ABB RAPID module: Ingenieria165.mod

MODULE Ingenieria165
    !***********************************************************
    !
    ! Modulo:  Ingenieria165
    !
    ! Descripción:
    !   Modulo con rutinas para decoracion con el motivo 165 años de facultad de ingeneria
    !
    ! Autor: Juan_Daleman
    !
    ! Versión: 1.0
    !
    !***********************************************************
    CONST robtarget Target_Tap165_10:=[[81.313,-88.677,-19.266],[0.707106781,0,0,0.707106781],[0,0,0,0],[9E+09,9E+09,9E+09,9E+09,9E+09,9E+09]];
    CONST robtarget Target_Tap165_20:=[[81.313,-88.677,-2.266],[0.707106781,0,0,0.707106781],[0,0,0,0],[9E+09,9E+09,9E+09,9E+09,9E+09,9E+09]];
    CONST robtarget Target_Tap165_30:=[[81.338,-82.631,-2.266],[0.707106781,0,0,0.707106781],[0,0,0,0],[9E+09,9E+09,9E+09,9E+09,9E+09,9E+09]];
    CONST robtarget Target_Tap165_40:=[[76.897,-82.904,-2.306],[0.707106781,0,0,0.707106781],[0,0,0,0],[9E+09,9E+09,9E+09,9E+09,9E+09,9E+09]];
    CONST robtarget Target_Tap165_50:=[[81.369,-82.46,-2.266],[0.707106781,0,0,0.707106781],[0,0,0,0],[9E+09,9E+09,9E+09,9E+09,9E+09,9E+09]];
    CONST robtarget Target_Tap165_60:=[[81.524,-77.183,-2.264],[0.707106781,0,0,0.707106781],[0,0,0,0],[9E+09,9E+09,9E+09,9E+09,9E+09,9E+09]];
    CONST robtarget Target_Tap165_70:=[[75.87,-77.461,-2.316],[0.707106781,0,0,0.707106781],[0,0,0,0],[9E+09,9E+09,9E+09,9E+09,9E+09,9E+09]];
    CONST robtarget Target_Tap165_80:=[[75.87,-77.461,-20],[0.707106781,0,0,0.707106781],[0,0,0,0],[9E+09,9E+09,9E+09,9E+09,9E+09,9E+09]];
    CONST robtarget Target_Tap165_90:=[[67.923,-79.66,-20],[0.707106781,0,0,0.707106781],[0,0,0,0],[9E+09,9E+09,9E+09,9E+09,9E+09,9E+09]];
    CONST robtarget Target_Tap165_100:=[[67.923,-79.66,-2.388],[0.707106781,0,0,0.707106781],[0,0,0,0],[9E+09,9E+09,9E+09,9E+09,9E+09,9E+09]];
    CONST robtarget Target_Tap165_110:=[[67.877,-88.682,-2.388],[0.707106781,0,0,0.707106781],[0,0,0,0],[9E+09,9E+09,9E+09,9E+09,9E+09,9E+09]];
    CONST robtarget Target_Tap165_120:=[[69.176,-87.545,-2.376],[0.707106781,0,0,0.707106781],[0,0,0,0],[9E+09,9E+09,9E+09,9E+09,9E+09,9E+09]];
    CONST robtarget Target_Tap165_130:=[[73.466,-88.301,-2.338],[0.707106781,0,0,0.707106781],[0,0,0,0],[9E+09,9E+09,9E+09,9E+09,9E+09,9E+09]];
    CONST robtarget Target_Tap165_140:=[[75.281,-84.884,-2.321],[0.707106781,0,0,0.707106781],[0,0,0,0],[9E+09,9E+09,9E+09,9E+09,9E+09,9E+09]];
    CONST robtarget Target_Tap165_150:=[[72.745,-79.717,-2.344],[0.707106781,0,0,0.707106781],[0,0,0,0],[9E+09,9E+09,9E+09,9E+09,9E+09,9E+09]];
    CONST robtarget Target_Tap165_160:=[[69.243,-80.87,-2.376],[0.707106781,0,0,0.707106781],[0,0,0,0],[9E+09,9E+09,9E+09,9E+09,9E+09,9E+09]];
    CONST robtarget Target_Tap165_170:=[[69.243,-80.87,-20],[0.707106781,0,0,0.707106781],[0,0,0,0],[9E+09,9E+09,9E+09,9E+09,9E+09,9E+09]];
    CONST robtarget Target_Tap165_180:=[[57.703,-85.818,-20],[0.707106781,0,0,0.707106781],[0,0,0,0],[9E+09,9E+09,9E+09,9E+09,9E+09,9E+09]];
    CONST robtarget Target_Tap165_190:=[[57.683,-85.747,-2.481],[0.707106781,0,0,0.707106781],[0,0,0,0],[9E+09,9E+09,9E+09,9E+09,9E+09,9E+09]];
    CONST robtarget Target_Tap165_200:=[[62.028,-88.896,-2.441],[0.707106781,0,0,0.707106781],[0,0,0,0],[9E+09,9E+09,9E+09,9E+09,9E+09,9E+09]];
    CONST robtarget Target_Tap165_210:=[[65.482,-83.568,-2.41],[0.707106781,0,0,0.707106781],[0,0,0,0],[9E+09,9E+09,9E+09,9E+09,9E+09,9E+09]];
    CONST robtarget Target_Tap165_220:=[[61.822,-79.686,-2.443],[0.707106781,0,0,0.707106781],[0,0,0,0],[9E+09,9E+09,9E+09,9E+09,9E+09,9E+09]];
    CONST robtarget Target_Tap165_230:=[[57.626,-82.905,-2.481],[0.707106781,0,0,0.707106781],[0,0,0,0],[9E+09,9E+09,9E+09,9E+09,9E+09,9E+09]];
    CONST robtarget Target_Tap165_240:=[[57.626,-82.905,-20],[0.707106781,0,0,0.707106781],[0,0,0,0],[9E+09,9E+09,9E+09,9E+09,9E+09,9E+09]];
    CONST robtarget Target_Tap165_250:=[[55.482,-79.946,-20],[0.707106781,0,0,0.707106781],[0,0,0,0],[9E+09,9E+09,9E+09,9E+09,9E+09,9E+09]];
    CONST robtarget Target_Tap165_260:=[[55.542,-79.789,-2.5],[0.707106781,0,0,0.707106781],[0,0,0,0],[9E+09,9E+09,9E+09,9E+09,9E+09,9E+09]];
    CONST robtarget Target_Tap165_270:=[[55.414,-88.257,-2.501],[0.707106781,0,0,0.707106781],[0,0,0,0],[9E+09,9E+09,9E+09,9E+09,9E+09,9E+09]];
    CONST robtarget Target_Tap165_280:=[[53.088,-88.957,-2.522],[0.707106781,0,0,0.707106781],[0,0,0,0],[9E+09,9E+09,9E+09,9E+09,9E+09,9E+09]];
    CONST robtarget Target_Tap165_290:=[[50.869,-87.673,-2.542],[0.707106781,0,0,0.707106781],[0,0,0,0],[9E+09,9E+09,9E+09,9E+09,9E+09,9E+09]];
    CONST robtarget Target_Tap165_300:=[[49.455,-88.876,-2.555],[0.707106781,0,0,0.707106781],[0,0,0,0],[9E+09,9E+09,9E+09,9E+09,9E+09,9E+09]];
    CONST robtarget Target_Tap165_310:=[[49.666,-79.854,-2.553],[0.707106781,0,0,0.707106781],[0,0,0,0],[9E+09,9E+09,9E+09,9E+09,9E+09,9E+09]];
    CONST robtarget Target_Tap165_320:=[[49.666,-79.854,-20],[0.707106781,0,0,0.707106781],[0,0,0,0],[9E+09,9E+09,9E+09,9E+09,9E+09,9E+09]];
    CONST robtarget Target_Tap165_330:=[[45.617,-88.918,-20],[0.707106781,0,0,0.707106781],[0,0,0,0],[9E+09,9E+09,9E+09,9E+09,9E+09,9E+09]];
    CONST robtarget Target_Tap165_340:=[[45.617,-88.918,-2.59],[0.707106781,0,0,0.707106781],[0,0,0,0],[9E+09,9E+09,9E+09,9E+09,9E+09,9E+09]];
    CONST robtarget Target_Tap165_350:=[[45.551,-76.897,-2.591],[0.707106781,0,0,0.707106781],[0,0,0,0],[9E+09,9E+09,9E+09,9E+09,9E+09,9E+09]];
    CONST robtarget Target_Tap165_360:=[[45.551,-76.897,-23],[0.707106781,0,0,0.707106781],[0,0,0,0],[9E+09,9E+09,9E+09,9E+09,9E+09,9E+09]];
    CONST robtarget Target_Tap165_370:=[[41.407,-77.76,-20],[0.707106781,0,0,0.707106781],[0,0,0,0],[9E+09,9E+09,9E+09,9E+09,9E+09,9E+09]];
    CONST robtarget Target_Tap165_380:=[[41.407,-77.76,0.372],[0.707106781,0,0,0.707106781],[0,0,0,0],[9E+09,9E+09,9E+09,9E+09,9E+09,9E+09]];
    CONST robtarget Target_Tap165_390:=[[41.282,-80.994,-2.629],[0.707106781,0,0,0.707106781],[0,0,0,0],[9E+09,9E+09,9E+09,9E+09,9E+09,9E+09]];
    CONST robtarget Target_Tap165_400:=[[43.422,-80.77,-2.61],[0.707106781,0,0,0.707106781],[0,0,0,0],[9E+09,9E+09,9E+09,9E+09,9E+09,9E+09]];
    CONST robtarget Target_Tap165_410:=[[38.361,-80.952,-2.656],[0.707106781,0,0,0.707106781],[0,0,0,0],[9E+09,9E+09,9E+09,9E+09,9E+09,9E+09]];
    CONST robtarget Target_Tap165_420:=[[41.333,-81.008,-2.629],[0.707106781,0,0,0.707106781],[0,0,0,0],[9E+09,9E+09,9E+09,9E+09,9E+09,9E+09]];
    CONST robtarget Target_Tap165_430:=[[41.267,-88.487,-2.629],[0.707106781,0,0,0.707106781],[0,0,0,0],[9E+09,9E+09,9E+09,9E+09,9E+09,9E+09]];
    CONST robtarget Target_Tap165_440:=[[38.45,-88.997,-2.655],[0.707106781,0,0,0.707106781],[0,0,0,0],[9E+09,9E+09,9E+09,9E+09,9E+09,9E+09]];
    CONST robtarget Target_Tap165_450:=[[38.45,-88.997,-20],[0.707106781,0,0,0.707106781],[0,0,0,0],[9E+09,9E+09,9E+09,9E+09,9E+09,9E+09]];
    CONST robtarget Target_Tap165_460:=[[30.389,-80.073,-20],[0.707106781,0,0,0.707106781],[0,0,0,0],[9E+09,9E+09,9E+09,9E+09,9E+09,9E+09]];
    CONST robtarget Target_Tap165_470:=[[30.389,-80.073,-2.728],[0.707106781,0,0,0.707106781],[0,0,0,0],[9E+09,9E+09,9E+09,9E+09,9E+09,9E+09]];
    CONST robtarget Target_Tap165_480:=[[30.235,-89.097,-2.73],[0.707106781,0,0,0.707106781],[0,0,0,0],[9E+09,9E+09,9E+09,9E+09,9E+09,9E+09]];
    CONST robtarget Target_Tap165_490:=[[31.518,-87.896,-2.718],[0.707106781,0,0,0.707106781],[0,0,0,0],[9E+09,9E+09,9E+09,9E+09,9E+09,9E+09]];
    CONST robtarget Target_Tap165_500:=[[34.632,-89.19,-2.69],[0.707106781,0,0,0.707106781],[0,0,0,0],[9E+09,9E+09,9E+09,9E+09,9E+09,9E+09]];
    CONST robtarget Target_Tap165_510:=[[37.622,-85.047,-2.663],[0.707106781,0,0,0.707106781],[0,0,0,0],[9E+09,9E+09,9E+09,9E+09,9E+09,9E+09]];
    CONST robtarget Target_Tap165_520:=[[35.565,-79.921,-2.682],[0.707106781,0,0,0.707106781],[0,0,0,0],[9E+09,9E+09,9E+09,9E+09,9E+09,9E+09]];
    CONST robtarget Target_Tap165_530:=[[31.419,-81.282,-2.719],[0.707106781,0,0,0.707106781],[0,0,0,0],[9E+09,9E+09,9E+09,9E+09,9E+09,9E+09]];
    CONST robtarget Target_Tap165_540:=[[31.419,-81.282,-20],[0.707106781,0,0,0.707106781],[0,0,0,0],[9E+09,9E+09,9E+09,9E+09,9E+09,9E+09]];
    CONST robtarget Target_Tap165_550:=[[20.747,-77.17,-20],[0.707106781,0,0,0.707106781],[0,0,0,0],[9E+09,9E+09,9E+09,9E+09,9E+09,9E+09]];
    CONST robtarget Target_Tap165_560:=[[20.805,-77.169,-2.815],[0.707106781,0,0,0.707106781],[0,0,0,0],[9E+09,9E+09,9E+09,9E+09,9E+09,9E+09]];
    CONST robtarget Target_Tap165_570:=[[20.61,-89.193,-2.817],[0.707106781,0,0,0.707106781],[0,0,0,0],[9E+09,9E+09,9E+09,9E+09,9E+09,9E+09]];
    CONST robtarget Target_Tap165_580:=[[21.819,-88.233,-2.806],[0.707106781,0,0,0.707106781],[0,0,0,0],[9E+09,9E+09,9E+09,9E+09,9E+09,9E+09]];
    CONST robtarget Target_Tap165_590:=[[25.21,-89.217,-2.775],[0.707106781,0,0,0.707106781],[0,0,0,0],[9E+09,9E+09,9E+09,9E+09,9E+09,9E+09]];
    CONST robtarget Target_Tap165_600:=[[27.949,-85.408,-2.75],[0.707106781,0,0,0.707106781],[0,0,0,0],[9E+09,9E+09,9E+09,9E+09,9E+09,9E+09]];
    CONST robtarget Target_Tap165_610:=[[25.874,-80.415,-2.769],[0.707106781,0,0,0.707106781],[0,0,0,0],[9E+09,9E+09,9E+09,9E+09,9E+09,9E+09]];
    CONST robtarget Target_Tap165_620:=[[21.748,-81.419,-2.807],[0.707106781,0,0,0.707106781],[0,0,0,0],[9E+09,9E+09,9E+09,9E+09,9E+09,9E+09]];
    CONST robtarget Target_Tap165_630:=[[21.748,-81.419,-20],[0.707106781,0,0,0.707106781],[0,0,0,0],[9E+09,9E+09,9E+09,9E+09,9E+09,9E+09]];
    CONST robtarget Target_Tap165_640:=[[8.35,-77.306,-20],[0.707106781,0,0,0.707106781],[0,0,0,0],[9E+09,9E+09,9E+09,9E+09,9E+09,9E+09]];
    CONST robtarget Target_Tap165_650:=[[8.35,-77.306,-2.928],[0.707106781,0,0,0.707106781],[0,0,0,0],[9E+09,9E+09,9E+09,9E+09,9E+09,9E+09]];
    CONST robtarget Target_Tap165_660:=[[7.975,-89.332,-2.932],[0.707106781,0,0,0.707106781],[0,0,0,0],[9E+09,9E+09,9E+09,9E+09,9E+09,9E+09]];
    CONST robtarget Target_Tap165_670:=[[9.494,-88.106,-2.918],[0.707106781,0,0,0.707106781],[0,0,0,0],[9E+09,9E+09,9E+09,9E+09,9E+09,9E+09]];
    CONST robtarget Target_Tap165_680:=[[13.081,-89.294,-2.885],[0.707106781,0,0,0.707106781],[0,0,0,0],[9E+09,9E+09,9E+09,9E+09,9E+09,9E+09]];
    CONST robtarget Target_Tap165_690:=[[15.593,-85.146,-2.863],[0.707106781,0,0,0.707106781],[0,0,0,0],[9E+09,9E+09,9E+09,9E+09,9E+09,9E+09]];
    CONST robtarget Target_Tap165_700:=[[13.446,-80.526,-2.882],[0.707106781,0,0,0.707106781],[0,0,0,0],[9E+09,9E+09,9E+09,9E+09,9E+09,9E+09]];
    CONST robtarget Target_Tap165_710:=[[9.38,-81.539,-2.919],[0.707106781,0,0,0.707106781],[0,0,0,0],[9E+09,9E+09,9E+09,9E+09,9E+09,9E+09]];
    CONST robtarget Target_Tap165_720:=[[9.38,-81.539,-20],[0.707106781,0,0,0.707106781],[0,0,0,0],[9E+09,9E+09,9E+09,9E+09,9E+09,9E+09]];
    CONST robtarget Target_Tap165_730:=[[-2.035,-86.612,-20],[0.707106781,0,0,0.707106781],[0,0,0,0],[9E+09,9E+09,9E+09,9E+09,9E+09,9E+09]];
    CONST robtarget Target_Tap165_740:=[[-2.035,-86.612,-3.023],[0.707106781,0,0,0.707106781],[0,0,0,0],[9E+09,9E+09,9E+09,9E+09,9E+09,9E+09]];
    CONST robtarget Target_Tap165_750:=[[2.246,-89.541,-2.984],[0.707106781,0,0,0.707106781],[0,0,0,0],[9E+09,9E+09,9E+09,9E+09,9E+09,9E+09]];
    CONST robtarget Target_Tap165_760:=[[5.81,-84.927,-2.951],[0.707106781,0,0,0.707106781],[0,0,0,0],[9E+09,9E+09,9E+09,9E+09,9E+09,9E+09]];
    CONST robtarget Target_Tap165_770:=[[1.692,-80.318,-2.989],[0.707106781,0,0,0.707106781],[0,0,0,0],[9E+09,9E+09,9E+09,9E+09,9E+09,9E+09]];
    CONST robtarget Target_Tap165_780:=[[-2.242,-85.619,-3.024],[0.707106781,0,0,0.707106781],[0,0,0,0],[9E+09,9E+09,9E+09,9E+09,9E+09,9E+09]];
    CONST robtarget Target_Tap165_790:=[[3.474,-85.692,-2.973],[0.707106781,0,0,0.707106781],[0,0,0,0],[9E+09,9E+09,9E+09,9E+09,9E+09,9E+09]];
    CONST robtarget Target_Tap165_800:=[[3.474,-85.692,-20],[0.707106781,0,0,0.707106781],[0,0,0,0],[9E+09,9E+09,9E+09,9E+09,9E+09,9E+09]];
    CONST robtarget Target_Tap165_810:=[[-7.455,-89.529,-20],[0.707106781,0,0,0.707106781],[0,0,0,0],[9E+09,9E+09,9E+09,9E+09,9E+09,9E+09]];
    CONST robtarget Target_Tap165_820:=[[-7.455,-89.529,-3.072],[0.707106781,0,0,0.707106781],[0,0,0,0],[9E+09,9E+09,9E+09,9E+09,9E+09,9E+09]];
    CONST robtarget Target_Tap165_830:=[[-7.408,-78.16,-3.071],[0.707106781,0,0,0.707106781],[0,0,0,0],[9E+09,9E+09,9E+09,9E+09,9E+09,9E+09]];
    CONST robtarget Target_Tap165_840:=[[-7.408,-78.16,-20],[0.707106781,0,0,0.707106781],[0,0,0,0],[9E+09,9E+09,9E+09,9E+09,9E+09,9E+09]];
    CONST robtarget Target_Tap165_850:=[[-11.373,-89.538,-20],[0.707106781,0,0,0.707106781],[0,0,0,0],[9E+09,9E+09,9E+09,9E+09,9E+09,9E+09]];
    CONST robtarget Target_Tap165_860:=[[-11.373,-89.538,-3.107],[0.707106781,0,0,0.707106781],[0,0,0,0],[9E+09,9E+09,9E+09,9E+09,9E+09,9E+09]];
    CONST robtarget Target_Tap165_870:=[[-11.145,-80.51,-3.105],[0.707106781,0,0,0.707106781],[0,0,0,0],[9E+09,9E+09,9E+09,9E+09,9E+09,9E+09]];
    CONST robtarget Target_Tap165_880:=[[-12.596,-81.788,-3.118],[0.707106781,0,0,0.707106781],[0,0,0,0],[9E+09,9E+09,9E+09,9E+09,9E+09,9E+09]];
    CONST robtarget Target_Tap165_890:=[[-15.49,-80.547,-3.145],[0.707106781,0,0,0.707106781],[0,0,0,0],[9E+09,9E+09,9E+09,9E+09,9E+09,9E+09]];
    CONST robtarget Target_Tap165_900:=[[-18.209,-83.364,-3.169],[0.707106781,0,0,0.707106781],[0,0,0,0],[9E+09,9E+09,9E+09,9E+09,9E+09,9E+09]];
    CONST robtarget Target_Tap165_910:=[[-18.164,-89.619,-3.169],[0.707106781,0,0,0.707106781],[0,0,0,0],[9E+09,9E+09,9E+09,9E+09,9E+09,9E+09]];
    CONST robtarget Target_Tap165_920:=[[-18.164,-89.619,-20],[0.707106781,0,0,0.707106781],[0,0,0,0],[9E+09,9E+09,9E+09,9E+09,9E+09,9E+09]];
    CONST robtarget Target_Tap165_930:=[[-19.664,-90.875,-20],[0.707106781,0,0,0.707106781],[0,0,0,0],[9E+09,9E+09,9E+09,9E+09,9E+09,9E+09]];
    CONST robtarget Target_Tap165_940:=[[-19.664,-90.875,-3.183],[0.707106781,0,0,0.707106781],[0,0,0,0],[9E+09,9E+09,9E+09,9E+09,9E+09,9E+09]];
    CONST robtarget Target_Tap165_950:=[[-24.113,-94.259,-3.223],[0.707106781,0,0,0.707106781],[0,0,0,0],[9E+09,9E+09,9E+09,9E+09,9E+09,9E+09]];
    CONST robtarget Target_Tap165_960:=[[-27.791,-90.884,-3.256],[0.707106781,0,0,0.707106781],[0,0,0,0],[9E+09,9E+09,9E+09,9E+09,9E+09,9E+09]];
    CONST robtarget Target_Tap165_970:=[[-27.929,-80.7,-3.258],[0.707106781,0,0,0.707106781],[0,0,0,0],[9E+09,9E+09,9E+09,9E+09,9E+09,9E+09]];
    CONST robtarget Target_Tap165_980:=[[-25.441,-81.899,-3.235],[0.707106781,0,0,0.707106781],[0,0,0,0],[9E+09,9E+09,9E+09,9E+09,9E+09,9E+09]];
    CONST robtarget Target_Tap165_990:=[[-22.502,-80.601,-3.208],[0.707106781,0,0,0.707106781],[0,0,0,0],[9E+09,9E+09,9E+09,9E+09,9E+09,9E+09]];
    CONST robtarget Target_Tap165_1000:=[[-19.387,-85.991,-3.18],[0.707106781,0,0,0.707106781],[0,0,0,0],[9E+09,9E+09,9E+09,9E+09,9E+09,9E+09]];
    CONST robtarget Target_Tap165_1010:=[[-21.158,-89.313,-3.196],[0.707106781,0,0,0.707106781],[0,0,0,0],[9E+09,9E+09,9E+09,9E+09,9E+09,9E+09]];
    CONST robtarget Target_Tap165_1020:=[[-25.481,-88.527,-3.235],[0.707106781,0,0,0.707106781],[0,0,0,0],[9E+09,9E+09,9E+09,9E+09,9E+09,9E+09]];
    CONST robtarget Target_Tap165_1030:=[[-25.431,-88.495,-20],[0.707106781,0,0,0.707106781],[0,0,0,0],[9E+09,9E+09,9E+09,9E+09,9E+09,9E+09]];
    CONST robtarget Target_Tap165_1040:=[[-36.83,-87.065,-20],[0.707106781,0,0,0.707106781],[0,0,0,0],[9E+09,9E+09,9E+09,9E+09,9E+09,9E+09]];
    CONST robtarget Target_Tap165_1050:=[[-36.83,-87.065,-3.338],[0.707106781,0,0,0.707106781],[0,0,0,0],[9E+09,9E+09,9E+09,9E+09,9E+09,9E+09]];
    CONST robtarget Target_Tap165_1060:=[[-32.555,-89.922,-3.3],[0.707106781,0,0,0.707106781],[0,0,0,0],[9E+09,9E+09,9E+09,9E+09,9E+09,9E+09]];
    CONST robtarget Target_Tap165_1070:=[[-29.008,-85.405,-3.267],[0.707106781,0,0,0.707106781],[0,0,0,0],[9E+09,9E+09,9E+09,9E+09,9E+09,9E+09]];
    CONST robtarget Target_Tap165_1080:=[[-33.253,-80.703,-3.306],[0.707106781,0,0,0.707106781],[0,0,0,0],[9E+09,9E+09,9E+09,9E+09,9E+09,9E+09]];
    CONST robtarget Target_Tap165_1090:=[[-37.045,-86.192,-3.34],[0.707106781,0,0,0.707106781],[0,0,0,0],[9E+09,9E+09,9E+09,9E+09,9E+09,9E+09]];
    CONST robtarget Target_Tap165_1100:=[[-31.341,-85.939,-3.289],[0.707106781,0,0,0.707106781],[0,0,0,0],[9E+09,9E+09,9E+09,9E+09,9E+09,9E+09]];
    CONST robtarget Target_Tap165_1110:=[[-31.341,-85.939,-20],[0.707106781,0,0,0.707106781],[0,0,0,0],[9E+09,9E+09,9E+09,9E+09,9E+09,9E+09]];
    CONST robtarget Target_Tap165_1120:=[[-39.521,-89.847,-20],[0.707106781,0,0,0.707106781],[0,0,0,0],[9E+09,9E+09,9E+09,9E+09,9E+09,9E+09]];
    CONST robtarget Target_Tap165_1130:=[[-39.521,-89.847,-3.363],[0.707106781,0,0,0.707106781],[0,0,0,0],[9E+09,9E+09,9E+09,9E+09,9E+09,9E+09]];
    CONST robtarget Target_Tap165_1140:=[[-39.341,-80.799,-3.361],[0.707106781,0,0,0.707106781],[0,0,0,0],[9E+09,9E+09,9E+09,9E+09,9E+09,9E+09]];
    CONST robtarget Target_Tap165_1150:=[[-40.79,-82.023,-3.374],[0.707106781,0,0,0.707106781],[0,0,0,0],[9E+09,9E+09,9E+09,9E+09,9E+09,9E+09]];
    CONST robtarget Target_Tap165_1160:=[[-43.877,-80.891,-3.402],[0.707106781,0,0,0.707106781],[0,0,0,0],[9E+09,9E+09,9E+09,9E+09,9E+09,9E+09]];
    CONST robtarget Target_Tap165_1170:=[[-46.356,-83.847,-3.425],[0.707106781,0,0,0.707106781],[0,0,0,0],[9E+09,9E+09,9E+09,9E+09,9E+09,9E+09]];
    CONST robtarget Target_Tap165_1180:=[[-46.289,-89.929,-3.424],[0.707106781,0,0,0.707106781],[0,0,0,0],[9E+09,9E+09,9E+09,9E+09,9E+09,9E+09]];
    CONST robtarget Target_Tap165_1190:=[[-46.289,-89.929,-20],[0.707106781,0,0,0.707106781],[0,0,0,0],[9E+09,9E+09,9E+09,9E+09,9E+09,9E+09]];
    CONST robtarget Target_Tap165_1200:=[[-49.014,-89.958,-20],[0.707106781,0,0,0.707106781],[0,0,0,0],[9E+09,9E+09,9E+09,9E+09,9E+09,9E+09]];
    CONST robtarget Target_Tap165_1210:=[[-49.014,-89.958,-3.449],[0.707106781,0,0,0.707106781],[0,0,0,0],[9E+09,9E+09,9E+09,9E+09,9E+09,9E+09]];
    CONST robtarget Target_Tap165_1220:=[[-48.979,-81.092,-3.449],[0.707106781,0,0,0.707106781],[0,0,0,0],[9E+09,9E+09,9E+09,9E+09,9E+09,9E+09]];
    CONST robtarget Target_Tap165_1230:=[[-48.979,-81.092,-20],[0.707106781,0,0,0.707106781],[0,0,0,0],[9E+09,9E+09,9E+09,9E+09,9E+09,9E+09]];
    CONST robtarget Target_Tap165_1240:=[[-49.066,-76.978,-20],[0.707106781,0,0,0.707106781],[0,0,0,0],[9E+09,9E+09,9E+09,9E+09,9E+09,9E+09]];
    CONST robtarget Target_Tap165_1250:=[[-49.066,-76.978,-3.449],[0.707106781,0,0,0.707106781],[0,0,0,0],[9E+09,9E+09,9E+09,9E+09,9E+09,9E+09]];
    CONST robtarget Target_Tap165_1260:=[[-49.067,-76.978,-20],[0.707106781,0,0,0.707106781],[0,0,0,0],[9E+09,9E+09,9E+09,9E+09,9E+09,9E+09]];
    CONST robtarget Target_Tap165_1270:=[[-59.116,-87.342,-20],[0.707106781,0,0,0.707106781],[0,0,0,0],[9E+09,9E+09,9E+09,9E+09,9E+09,9E+09]];
    CONST robtarget Target_Tap165_1280:=[[-59.127,-87.309,-3.541],[0.707106781,0,0,0.707106781],[0,0,0,0],[9E+09,9E+09,9E+09,9E+09,9E+09,9E+09]];
    CONST robtarget Target_Tap165_1290:=[[-54.679,-90.143,-3.5],[0.707106781,0,0,0.707106781],[0,0,0,0],[9E+09,9E+09,9E+09,9E+09,9E+09,9E+09]];
    CONST robtarget Target_Tap165_1300:=[[-51.303,-85.577,-3.47],[0.707106781,0,0,0.707106781],[0,0,0,0],[9E+09,9E+09,9E+09,9E+09,9E+09,9E+09]];
    CONST robtarget Target_Tap165_1310:=[[-55.273,-80.95,-3.506],[0.707106781,0,0,0.707106781],[0,0,0,0],[9E+09,9E+09,9E+09,9E+09,9E+09,9E+09]];
    CONST robtarget Target_Tap165_1320:=[[-59.346,-86.247,-3.543],[0.707106781,0,0,0.707106781],[0,0,0,0],[9E+09,9E+09,9E+09,9E+09,9E+09,9E+09]];
    CONST robtarget Target_Tap165_1330:=[[-53.484,-85.871,-3.489],[0.707106781,0,0,0.707106781],[0,0,0,0],[9E+09,9E+09,9E+09,9E+09,9E+09,9E+09]];
    CONST robtarget Target_Tap165_1340:=[[-53.484,-85.871,-20],[0.707106781,0,0,0.707106781],[0,0,0,0],[9E+09,9E+09,9E+09,9E+09,9E+09,9E+09]];
    CONST robtarget Target_Tap165_1350:=[[-61.947,-90.17,-20],[0.707106781,0,0,0.707106781],[0,0,0,0],[9E+09,9E+09,9E+09,9E+09,9E+09,9E+09]];
    CONST robtarget Target_Tap165_1360:=[[-61.843,-89.868,-3.565],[0.707106781,0,0,0.707106781],[0,0,0,0],[9E+09,9E+09,9E+09,9E+09,9E+09,9E+09]];
    CONST robtarget Target_Tap165_1370:=[[-61.597,-81.121,-3.563],[0.707106781,0,0,0.707106781],[0,0,0,0],[9E+09,9E+09,9E+09,9E+09,9E+09,9E+09]];
    CONST robtarget Target_Tap165_1380:=[[-62.926,-82.842,-3.575],[0.707106781,0,0,0.707106781],[0,0,0,0],[9E+09,9E+09,9E+09,9E+09,9E+09,9E+09]];
    CONST robtarget Target_Tap165_1390:=[[-65.595,-81.119,-3.599],[0.707106781,0,0,0.707106781],[0,0,0,0],[9E+09,9E+09,9E+09,9E+09,9E+09,9E+09]];
    CONST robtarget Target_Tap165_1400:=[[-65.595,-81.119,-20],[0.707106781,0,0,0.707106781],[0,0,0,0],[9E+09,9E+09,9E+09,9E+09,9E+09,9E+09]];
    CONST robtarget Target_Tap165_1410:=[[-66.223,-79.394,-20],[0.707106781,0,0,0.707106781],[0,0,0,0],[9E+09,9E+09,9E+09,9E+09,9E+09,9E+09]];
    CONST robtarget Target_Tap165_1420:=[[-66.223,-79.394,-3.605],[0.707106781,0,0,0.707106781],[0,0,0,0],[9E+09,9E+09,9E+09,9E+09,9E+09,9E+09]];
    CONST robtarget Target_Tap165_1430:=[[-69.594,-77.785,-3.636],[0.707106781,0,0,0.707106781],[0,0,0,0],[9E+09,9E+09,9E+09,9E+09,9E+09,9E+09]];
    CONST robtarget Target_Tap165_1440:=[[-69.594,-77.785,-20],[0.707106781,0,0,0.707106781],[0,0,0,0],[9E+09,9E+09,9E+09,9E+09,9E+09,9E+09]];
    CONST robtarget Target_Tap165_1450:=[[-67.838,-81.282,-20],[0.707106781,0,0,0.707106781],[0,0,0,0],[9E+09,9E+09,9E+09,9E+09,9E+09,9E+09]];
    CONST robtarget Target_Tap165_1460:=[[-67.838,-81.282,-3.62],[0.707106781,0,0,0.707106781],[0,0,0,0],[9E+09,9E+09,9E+09,9E+09,9E+09,9E+09]];
    CONST robtarget Target_Tap165_1470:=[[-67.868,-90.166,-3.62],[0.707106781,0,0,0.707106781],[0,0,0,0],[9E+09,9E+09,9E+09,9E+09,9E+09,9E+09]];
    CONST robtarget Target_Tap165_1480:=[[-67.868,-90.166,-20.62],[0.707106781,0,0,0.707106781],[0,0,0,0],[9E+09,9E+09,9E+09,9E+09,9E+09,9E+09]];
    CONST robtarget Target_Tap165_1490:=[[-77.715,-81.363,-20],[0.707106781,0,0,0.707106781],[0,0,0,0],[9E+09,9E+09,9E+09,9E+09,9E+09,9E+09]];
    CONST robtarget Target_Tap165_1500:=[[-77.715,-81.363,-3.709],[0.707106781,0,0,0.707106781],[0,0,0,0],[9E+09,9E+09,9E+09,9E+09,9E+09,9E+09]];
    CONST robtarget Target_Tap165_1510:=[[-78.085,-90.282,-3.713],[0.707106781,0,0,0.707106781],[0,0,0,0],[9E+09,9E+09,9E+09,9E+09,9E+09,9E+09]];
    CONST robtarget Target_Tap165_1520:=[[-76.677,-89.371,-3.7],[0.707106781,0,0,0.707106781],[0,0,0,0],[9E+09,9E+09,9E+09,9E+09,9E+09,9E+09]];
    CONST robtarget Target_Tap165_1530:=[[-72.593,-90.069,-3.663],[0.707106781,0,0,0.707106781],[0,0,0,0],[9E+09,9E+09,9E+09,9E+09,9E+09,9E+09]];
    CONST robtarget Target_Tap165_1540:=[[-70.623,-84.883,-3.645],[0.707106781,0,0,0.707106781],[0,0,0,0],[9E+09,9E+09,9E+09,9E+09,9E+09,9E+09]];
    CONST robtarget Target_Tap165_1550:=[[-74.575,-81.203,-3.681],[0.707106781,0,0,0.707106781],[0,0,0,0],[9E+09,9E+09,9E+09,9E+09,9E+09,9E+09]];
    CONST robtarget Target_Tap165_1560:=[[-76.614,-82.474,-3.699],[0.707106781,0,0,0.707106781],[0,0,0,0],[9E+09,9E+09,9E+09,9E+09,9E+09,9E+09]];
    CONST robtarget Target_Tap165_1570:=[[-76.614,-82.474,-20],[0.707106781,0,0,0.707106781],[0,0,0,0],[9E+09,9E+09,9E+09,9E+09,9E+09,9E+09]];
    CONST robtarget Target_Tap165_1580:=[[-39.17,-32.252,-20],[0.707106781,0,0,0.707106781],[0,-1,0,0],[9E+09,9E+09,9E+09,9E+09,9E+09,9E+09]];
    CONST robtarget Target_Tap165_1590:=[[-39.17,-32.252,-3.36],[0.707106781,0,0,0.707106781],[0,-1,0,0],[9E+09,9E+09,9E+09,9E+09,9E+09,9E+09]];
    CONST robtarget Target_Tap165_1600:=[[-45.406,-40.686,-3.416],[0.707106781,0,0,0.707106781],[0,-1,0,0],[9E+09,9E+09,9E+09,9E+09,9E+09,9E+09]];
    CONST robtarget Target_Tap165_1610:=[[-56.317,-45.81,-3.515],[0.707106781,0,0,0.707106781],[0,-1,0,0],[9E+09,9E+09,9E+09,9E+09,9E+09,9E+09]];
    CONST robtarget Target_Tap165_1620:=[[-56.318,-45.719,-20],[0.707106781,0,0,0.707106781],[0,-1,0,0],[9E+09,9E+09,9E+09,9E+09,9E+09,9E+09]];
    CONST robtarget Target_Tap165_1630:=[[-59.302,-45.926,-20],[0.707106781,0,0,0.707106781],[0,-1,0,0],[9E+09,9E+09,9E+09,9E+09,9E+09,9E+09]];
    CONST robtarget Target_Tap165_1640:=[[-59.302,-45.926,-2.542],[0.707106781,0,0,0.707106781],[0,-1,0,0],[9E+09,9E+09,9E+09,9E+09,9E+09,9E+09]];
    CONST robtarget Target_Tap165_1650:=[[-71.823,-39.415,-2.656],[0.707106781,0,0,0.707106781],[0,-1,0,0],[9E+09,9E+09,9E+09,9E+09,9E+09,9E+09]];
    CONST robtarget Target_Tap165_1660:=[[-78.717,-24.374,-2.719],[0.707106781,0,0,0.707106781],[0,-1,0,0],[9E+09,9E+09,9E+09,9E+09,9E+09,9E+09]];
    CONST robtarget Target_Tap165_1670:=[[-78.717,-24.374,-20],[0.707106781,0,0,0.707106781],[0,-1,0,0],[9E+09,9E+09,9E+09,9E+09,9E+09,9E+09]];
    CONST robtarget Target_Tap165_1680:=[[-78.807,-20.649,-20],[0.707106781,0,0,0.707106781],[0,-1,0,0],[9E+09,9E+09,9E+09,9E+09,9E+09,9E+09]];
    CONST robtarget Target_Tap165_1690:=[[-78.607,-20.647,-2.718],[0.707106781,0,0,0.707106781],[0,-1,0,0],[9E+09,9E+09,9E+09,9E+09,9E+09,9E+09]];
    CONST robtarget Target_Tap165_1700:=[[-72.81,-6.435,-2.665],[0.707106781,0,0,0.707106781],[0,-1,0,0],[9E+09,9E+09,9E+09,9E+09,9E+09,9E+09]];
    CONST robtarget Target_Tap165_1710:=[[-59.701,1.288,-2.546],[0.707106781,0,0,0.707106781],[0,-1,0,0],[9E+09,9E+09,9E+09,9E+09,9E+09,9E+09]];
    CONST robtarget Target_Tap165_1720:=[[-59.701,1.288,-20],[0.707106781,0,0,0.707106781],[0,-1,0,0],[9E+09,9E+09,9E+09,9E+09,9E+09,9E+09]];
    CONST robtarget Target_Tap165_1730:=[[-52.716,-4.037,-20],[0.707106781,0,0,0.707106781],[0,-1,0,0],[9E+09,9E+09,9E+09,9E+09,9E+09,9E+09]];
    CONST robtarget Target_Tap165_1740:=[[-52.716,-4.037,-2.483],[0.707106781,0,0,0.707106781],[0,-1,0,0],[9E+09,9E+09,9E+09,9E+09,9E+09,9E+09]];
    CONST robtarget Target_Tap165_1750:=[[-52.662,15.745,-2.482],[0.707106781,0,0,0.707106781],[0,0,0,0],[9E+09,9E+09,9E+09,9E+09,9E+09,9E+09]];
    CONST robtarget Target_Tap165_1760:=[[-52.662,15.745,-20],[0.707106781,0,0,0.707106781],[0,0,0,0],[9E+09,9E+09,9E+09,9E+09,9E+09,9E+09]];
    CONST robtarget Target_Tap165_1770:=[[-60.093,13.08,-20],[0.707106781,0,0,0.707106781],[0,0,0,0],[9E+09,9E+09,9E+09,9E+09,9E+09,9E+09]];
    CONST robtarget Target_Tap165_1780:=[[-60.065,13.257,-2.549],[0.707106781,0,0,0.707106781],[0,0,0,0],[9E+09,9E+09,9E+09,9E+09,9E+09,9E+09]];
    CONST robtarget Target_Tap165_1790:=[[-76.563,5.247,-2.699],[0.707106781,0,0,0.707106781],[0,0,0,0],[9E+09,9E+09,9E+09,9E+09,9E+09,9E+09]];
    CONST robtarget Target_Tap165_1800:=[[-89.184,-20.892,-2.814],[0.707106781,0,0,0.707106781],[0,0,0,0],[9E+09,9E+09,9E+09,9E+09,9E+09,9E+09]];
    CONST robtarget Target_Tap165_1810:=[[-89.184,-20.892,-20],[0.707106781,0,0,0.707106781],[0,0,0,0],[9E+09,9E+09,9E+09,9E+09,9E+09,9E+09]];
    CONST robtarget Target_Tap165_1820:=[[-89.283,-24.553,-20],[0.707106781,0,0,0.707106781],[0,0,0,0],[9E+09,9E+09,9E+09,9E+09,9E+09,9E+09]];
    CONST robtarget Target_Tap165_1830:=[[-89.283,-24.553,-3.814],[0.707106781,0,0,0.707106781],[0,0,0,0],[9E+09,9E+09,9E+09,9E+09,9E+09,9E+09]];
    CONST robtarget Target_Tap165_1840:=[[-79.776,-46.415,-3.728],[0.707106781,0,0,0.707106781],[0,0,0,0],[9E+09,9E+09,9E+09,9E+09,9E+09,9E+09]];
    CONST robtarget Target_Tap165_1850:=[[-59.333,-57.044,-3.542],[0.707106781,0,0,0.707106781],[0,0,0,0],[9E+09,9E+09,9E+09,9E+09,9E+09,9E+09]];
    CONST robtarget Target_Tap165_1860:=[[-59.333,-57.044,-20],[0.707106781,0,0,0.707106781],[0,0,0,0],[9E+09,9E+09,9E+09,9E+09,9E+09,9E+09]];
    CONST robtarget Target_Tap165_1870:=[[-56.192,-57.204,-20],[0.707106781,0,0,0.707106781],[0,0,0,0],[9E+09,9E+09,9E+09,9E+09,9E+09,9E+09]];
    CONST robtarget Target_Tap165_1880:=[[-56.192,-57.204,-3.514],[0.707106781,0,0,0.707106781],[0,0,0,0],[9E+09,9E+09,9E+09,9E+09,9E+09,9E+09]];
    CONST robtarget Target_Tap165_1890:=[[-37.634,-48.244,-3.346],[0.707106781,0,0,0.707106781],[0,0,0,0],[9E+09,9E+09,9E+09,9E+09,9E+09,9E+09]];
    CONST robtarget Target_Tap165_1900:=[[-28.695,-32.279,-3.265],[0.707106781,0,0,0.707106781],[0,0,0,0],[9E+09,9E+09,9E+09,9E+09,9E+09,9E+09]];
    CONST robtarget Target_Tap165_1910:=[[-28.695,-32.279,-20],[0.707106781,0,0,0.707106781],[0,0,0,0],[9E+09,9E+09,9E+09,9E+09,9E+09,9E+09]];
    CONST robtarget Target_Tap165_1920:=[[-31.717,-18.062,-20],[0.707106781,0,0,0.707106781],[0,0,0,0],[9E+09,9E+09,9E+09,9E+09,9E+09,9E+09]];
    CONST robtarget Target_Tap165_1930:=[[-31.717,-18.062,-3.292],[0.707106781,0,0,0.707106781],[0,0,0,0],[9E+09,9E+09,9E+09,9E+09,9E+09,9E+09]];
    CONST robtarget Target_Tap165_1940:=[[-31.82,-25.861,-3.293],[0.707106781,0,0,0.707106781],[0,0,0,0],[9E+09,9E+09,9E+09,9E+09,9E+09,9E+09]];
    CONST robtarget Target_Tap165_1950:=[[-30.999,-24.646,-3.285],[0.707106781,0,0,0.707106781],[0,0,0,0],[9E+09,9E+09,9E+09,9E+09,9E+09,9E+09]];
    CONST robtarget Target_Tap165_1960:=[[-28.081,-25.977,-3.259],[0.707106781,0,0,0.707106781],[0,0,0,0],[9E+09,9E+09,9E+09,9E+09,9E+09,9E+09]];
    CONST robtarget Target_Tap165_1970:=[[-25.106,-21.451,-3.232],[0.707106781,0,0,0.707106781],[0,0,0,0],[9E+09,9E+09,9E+09,9E+09,9E+09,9E+09]];
    CONST robtarget Target_Tap165_1980:=[[-27.038,-18.261,-3.25],[0.707106781,0,0,0.707106781],[0,0,0,0],[9E+09,9E+09,9E+09,9E+09,9E+09,9E+09]];
    CONST robtarget Target_Tap165_1990:=[[-31.054,-19.278,-3.286],[0.707106781,0,0,0.707106781],[0,0,0,0],[9E+09,9E+09,9E+09,9E+09,9E+09,9E+09]];
    CONST robtarget Target_Tap165_2000:=[[-31.054,-19.278,-20],[0.707106781,0,0,0.707106781],[0,0,0,0],[9E+09,9E+09,9E+09,9E+09,9E+09,9E+09]];
    CONST robtarget Target_Tap165_2010:=[[-35.765,-25.906,-20.329],[0.707106781,0,0,0.707106781],[0,0,0,0],[9E+09,9E+09,9E+09,9E+09,9E+09,9E+09]];
    CONST robtarget Target_Tap165_2020:=[[-35.765,-25.906,-3.329],[0.707106781,0,0,0.707106781],[0,0,0,0],[9E+09,9E+09,9E+09,9E+09,9E+09,9E+09]];
    CONST robtarget Target_Tap165_2030:=[[-35.772,-18.109,-3.329],[0.707106781,0,0,0.707106781],[0,0,0,0],[9E+09,9E+09,9E+09,9E+09,9E+09,9E+09]];
    CONST robtarget Target_Tap165_2040:=[[-36.461,-19.071,-3.335],[0.707106781,0,0,0.707106781],[0,0,0,0],[9E+09,9E+09,9E+09,9E+09,9E+09,9E+09]];
    CONST robtarget Target_Tap165_2050:=[[-38.585,-18.081,-3.354],[0.707106781,0,0,0.707106781],[0,0,0,0],[9E+09,9E+09,9E+09,9E+09,9E+09,9E+09]];
    CONST robtarget Target_Tap165_2060:=[[-41.065,-19.34,-3.377],[0.707106781,0,0,0.707106781],[0,0,0,0],[9E+09,9E+09,9E+09,9E+09,9E+09,9E+09]];
    CONST robtarget Target_Tap165_2070:=[[-41.588,-20.881,-3.382],[0.707106781,0,0,0.707106781],[0,0,0,0],[9E+09,9E+09,9E+09,9E+09,9E+09,9E+09]];
    CONST robtarget Target_Tap165_2080:=[[-41.405,-26,-3.38],[0.707106781,0,0,0.707106781],[0,0,0,0],[9E+09,9E+09,9E+09,9E+09,9E+09,9E+09]];
    CONST robtarget Target_Tap165_2090:=[[-41.405,-26,-20],[0.707106781,0,0,0.707106781],[0,0,0,0],[9E+09,9E+09,9E+09,9E+09,9E+09,9E+09]];
    CONST robtarget Target_Tap165_2100:=[[-36.486,-17.117,-20],[0.707106781,0,0,0.707106781],[0,0,0,0],[9E+09,9E+09,9E+09,9E+09,9E+09,9E+09]];
    CONST robtarget Target_Tap165_2110:=[[-36.53,-17.222,-3.336],[0.707106781,0,0,0.707106781],[0,0,0,0],[9E+09,9E+09,9E+09,9E+09,9E+09,9E+09]];
    CONST robtarget Target_Tap165_2120:=[[-37.445,-16.119,-3.344],[0.707106781,0,0,0.707106781],[0,0,0,0],[9E+09,9E+09,9E+09,9E+09,9E+09,9E+09]];
    CONST robtarget Target_Tap165_2130:=[[-38.411,-16.432,-3.353],[0.707106781,0,0,0.707106781],[0,0,0,0],[9E+09,9E+09,9E+09,9E+09,9E+09,9E+09]];
    CONST robtarget Target_Tap165_2140:=[[-39.286,-16.899,-3.361],[0.707106781,0,0,0.707106781],[0,0,0,0],[9E+09,9E+09,9E+09,9E+09,9E+09,9E+09]];
    CONST robtarget Target_Tap165_2150:=[[-40.378,-15.741,-3.371],[0.707106781,0,0,0.707106781],[0,0,0,0],[9E+09,9E+09,9E+09,9E+09,9E+09,9E+09]];
    CONST robtarget Target_Tap165_2160:=[[-40.386,-15.73,-20],[0.707106781,0,0,0.707106781],[0,0,0,0],[9E+09,9E+09,9E+09,9E+09,9E+09,9E+09]];
    CONST robtarget Target_Tap165_2170:=[[-47.314,-18.189,-20],[0.707106781,0,0,0.707106781],[0,0,0,0],[9E+09,9E+09,9E+09,9E+09,9E+09,9E+09]];
    CONST robtarget Target_Tap165_2180:=[[-47.314,-18.189,-3.434],[0.707106781,0,0,0.707106781],[0,0,0,0],[9E+09,9E+09,9E+09,9E+09,9E+09,9E+09]];
    CONST robtarget Target_Tap165_2190:=[[-51.125,-21.796,-3.468],[0.707106781,0,0,0.707106781],[0,0,0,0],[9E+09,9E+09,9E+09,9E+09,9E+09,9E+09]];
    CONST robtarget Target_Tap165_2200:=[[-47.362,-26.225,-3.434],[0.707106781,0,0,0.707106781],[0,0,0,0],[9E+09,9E+09,9E+09,9E+09,9E+09,9E+09]];
    CONST robtarget Target_Tap165_2210:=[[-43.935,-21.99,-3.403],[0.707106781,0,0,0.707106781],[0,0,0,0],[9E+09,9E+09,9E+09,9E+09,9E+09,9E+09]];
    CONST robtarget Target_Tap165_2220:=[[-47.266,-18.155,-3.433],[0.707106781,0,0,0.707106781],[0,0,0,0],[9E+09,9E+09,9E+09,9E+09,9E+09,9E+09]];
    CONST robtarget Target_Tap165_2230:=[[-47.266,-18.155,-20],[0.707106781,0,0,0.707106781],[0,0,0,0],[9E+09,9E+09,9E+09,9E+09,9E+09,9E+09]];
    CONST robtarget Target_Tap165_2240:=[[-57.971,-20.731,-20],[0.707106781,0,0,0.707106781],[0,0,0,0],[9E+09,9E+09,9E+09,9E+09,9E+09,9E+09]];
    CONST robtarget Target_Tap165_2250:=[[-57.971,-20.731,-3.53],[0.707106781,0,0,0.707106781],[0,0,0,0],[9E+09,9E+09,9E+09,9E+09,9E+09,9E+09]];
    CONST robtarget Target_Tap165_2260:=[[-55.993,-18.217,-3.512],[0.707106781,0,0,0.707106781],[0,0,0,0],[9E+09,9E+09,9E+09,9E+09,9E+09,9E+09]];
    CONST robtarget Target_Tap165_2270:=[[-53.238,-20.399,-3.487],[0.707106781,0,0,0.707106781],[0,0,0,0],[9E+09,9E+09,9E+09,9E+09,9E+09,9E+09]];
    CONST robtarget Target_Tap165_2280:=[[-53.464,-21.529,-3.489],[0.707106781,0,0,0.707106781],[0,0,0,0],[9E+09,9E+09,9E+09,9E+09,9E+09,9E+09]];
    CONST robtarget Target_Tap165_2290:=[[-58.489,-23.157,-3.535],[0.707106781,0,0,0.707106781],[0,0,0,0],[9E+09,9E+09,9E+09,9E+09,9E+09,9E+09]];
    CONST robtarget Target_Tap165_2300:=[[-55.943,-26.308,-3.512],[0.707106781,0,0,0.707106781],[0,0,0,0],[9E+09,9E+09,9E+09,9E+09,9E+09,9E+09]];
    CONST robtarget Target_Tap165_2310:=[[-53.104,-23.931,-3.486],[0.707106781,0,0,0.707106781],[0,0,0,0],[9E+09,9E+09,9E+09,9E+09,9E+09,9E+09]];
    CONST robtarget Target_Tap165_2320:=[[-53.104,-23.931,-20],[0.707106781,0,0,0.707106781],[0,0,0,0],[9E+09,9E+09,9E+09,9E+09,9E+09,9E+09]];
    CONST robtarget Target_Tap165_2330:=[[-41.125,31.366,-20],[0.707106781,0,0,0.707106781],[0,0,0,0],[9E+09,9E+09,9E+09,9E+09,9E+09,9E+09]];
    CONST robtarget Target_Tap165_2340:=[[-41.125,31.366,-3.377],[0.707106781,0,0,0.707106781],[0,0,0,0],[9E+09,9E+09,9E+09,9E+09,9E+09,9E+09]];
    CONST robtarget Target_Tap165_2350:=[[-40.788,-11.491,-3.374],[0.707106781,0,0,0.707106781],[0,0,0,0],[9E+09,9E+09,9E+09,9E+09,9E+09,9E+09]];
    CONST robtarget Target_Tap165_2360:=[[-40.788,-11.491,-20],[0.707106781,0,0,0.707106781],[0,0,0,0],[9E+09,9E+09,9E+09,9E+09,9E+09,9E+09]];
    CONST robtarget Target_Tap165_2370:=[[-30.616,-11.403,-20],[0.707106781,0,0,0.707106781],[0,0,0,0],[9E+09,9E+09,9E+09,9E+09,9E+09,9E+09]];
    CONST robtarget Target_Tap165_2380:=[[-30.616,-11.403,-3.282],[0.707106781,0,0,0.707106781],[0,0,0,0],[9E+09,9E+09,9E+09,9E+09,9E+09,9E+09]];
    CONST robtarget Target_Tap165_2390:=[[-30.714,31.592,-3.283],[0.707106781,0,0,0.707106781],[0,0,0,0],[9E+09,9E+09,9E+09,9E+09,9E+09,9E+09]];
    CONST robtarget Target_Tap165_2400:=[[-30.714,31.592,-20],[0.707106781,0,0,0.707106781],[0,0,0,0],[9E+09,9E+09,9E+09,9E+09,9E+09,9E+09]];
    CONST robtarget Target_Tap165_2410:=[[-27.739,39.945,-20],[0.707106781,0,0,0.707106781],[0,0,0,0],[9E+09,9E+09,9E+09,9E+09,9E+09,9E+09]];
    CONST robtarget Target_Tap165_2420:=[[-27.688,39.876,-2.255],[0.707106781,0,0,0.707106781],[0,0,0,0],[9E+09,9E+09,9E+09,9E+09,9E+09,9E+09]];
    CONST robtarget Target_Tap165_2430:=[[-86.73,38.296,-2.791],[0.707106781,0,0,0.707106781],[0,0,0,0],[9E+09,9E+09,9E+09,9E+09,9E+09,9E+09]];
    CONST robtarget Target_Tap165_2440:=[[-86.73,38.296,-20],[0.707106781,0,0,0.707106781],[0,0,0,0],[9E+09,9E+09,9E+09,9E+09,9E+09,9E+09]];
    CONST robtarget Target_Tap165_2450:=[[-86.961,50.097,-20],[0.707106781,0,0,0.707106781],[0,0,0,0],[9E+09,9E+09,9E+09,9E+09,9E+09,9E+09]];
    CONST robtarget Target_Tap165_2460:=[[-86.961,50.097,-2.793],[0.707106781,0,0,0.707106781],[0,0,0,0],[9E+09,9E+09,9E+09,9E+09,9E+09,9E+09]];
    CONST robtarget Target_Tap165_2470:=[[-27.534,50.96,-2.254],[0.707106781,0,0,0.707106781],[0,0,0,0],[9E+09,9E+09,9E+09,9E+09,9E+09,9E+09]];
    CONST robtarget Target_Tap165_2480:=[[-27.534,50.96,-20],[0.707106781,0,0,0.707106781],[0,0,0,0],[9E+09,9E+09,9E+09,9E+09,9E+09,9E+09]];
    CONST robtarget Target_Tap165_2490:=[[12.127,13.216,-20],[0.707106781,0,0,0.707106781],[0,0,0,0],[9E+09,9E+09,9E+09,9E+09,9E+09,9E+09]];
    CONST robtarget Target_Tap165_2500:=[[12.127,13.216,-2.894],[0.707106781,0,0,0.707106781],[0,0,0,0],[9E+09,9E+09,9E+09,9E+09,9E+09,9E+09]];
    CONST robtarget Target_Tap165_2510:=[[-8.993,1.151,-3.086],[0.707106781,0,0,0.707106781],[0,0,0,0],[9E+09,9E+09,9E+09,9E+09,9E+09,9E+09]];
    CONST robtarget Target_Tap165_2520:=[[-16.655,-19.965,-3.155],[0.707106781,0,0,0.707106781],[0,0,0,0],[9E+09,9E+09,9E+09,9E+09,9E+09,9E+09]];
    CONST robtarget Target_Tap165_2530:=[[-16.655,-19.965,-20],[0.707106781,0,0,0.707106781],[0,0,0,0],[9E+09,9E+09,9E+09,9E+09,9E+09,9E+09]];
    CONST robtarget Target_Tap165_2540:=[[-16.841,-23.499,-20],[0.707106781,0,0,0.707106781],[0,0,0,0],[9E+09,9E+09,9E+09,9E+09,9E+09,9E+09]];
    CONST robtarget Target_Tap165_2550:=[[-16.841,-23.499,-3.157],[0.707106781,0,0,0.707106781],[0,0,0,0],[9E+09,9E+09,9E+09,9E+09,9E+09,9E+09]];
    CONST robtarget Target_Tap165_2560:=[[-5.052,-48.573,-3.05],[0.707106781,0,0,0.707106781],[0,0,0,0],[9E+09,9E+09,9E+09,9E+09,9E+09,9E+09]];
    CONST robtarget Target_Tap165_2570:=[[13.646,-56.818,-2.88],[0.707106781,0,0,0.707106781],[0,0,0,0],[9E+09,9E+09,9E+09,9E+09,9E+09,9E+09]];
    CONST robtarget Target_Tap165_2580:=[[13.646,-56.818,-20],[0.707106781,0,0,0.707106781],[0,0,0,0],[9E+09,9E+09,9E+09,9E+09,9E+09,9E+09]];
    CONST robtarget Target_Tap165_2590:=[[16.904,-56.415,-20],[0.707106781,0,0,0.707106781],[0,0,0,0],[9E+09,9E+09,9E+09,9E+09,9E+09,9E+09]];
    CONST robtarget Target_Tap165_2600:=[[16.904,-56.415,-2.851],[0.707106781,0,0,0.707106781],[0,0,0,0],[9E+09,9E+09,9E+09,9E+09,9E+09,9E+09]];
    CONST robtarget Target_Tap165_2610:=[[37.054,-46.771,-2.668],[0.707106781,0,0,0.707106781],[0,0,0,0],[9E+09,9E+09,9E+09,9E+09,9E+09,9E+09]];
    CONST robtarget Target_Tap165_2620:=[[47.119,-22.803,-2.576],[0.707106781,0,0,0.707106781],[0,0,0,0],[9E+09,9E+09,9E+09,9E+09,9E+09,9E+09]];
    CONST robtarget Target_Tap165_2630:=[[47.119,-22.803,-20],[0.707106781,0,0,0.707106781],[0,0,0,0],[9E+09,9E+09,9E+09,9E+09,9E+09,9E+09]];
    CONST robtarget Target_Tap165_2640:=[[47.592,-19.252,-20],[0.707106781,0,0,0.707106781],[0,0,0,0],[9E+09,9E+09,9E+09,9E+09,9E+09,9E+09]];
    CONST robtarget Target_Tap165_2650:=[[47.592,-19.252,-2.572],[0.707106781,0,0,0.707106781],[0,0,0,0],[9E+09,9E+09,9E+09,9E+09,9E+09,9E+09]];
    CONST robtarget Target_Tap165_2660:=[[44.976,-9.049,-2.596],[0.707106781,0,0,0.707106781],[0,0,0,0],[9E+09,9E+09,9E+09,9E+09,9E+09,9E+09]];
    CONST robtarget Target_Tap165_2670:=[[43.625,-3.637,-2.608],[0.707106781,0,0,0.707106781],[0,0,0,0],[9E+09,9E+09,9E+09,9E+09,9E+09,9E+09]];
    CONST robtarget Target_Tap165_2680:=[[9.76,55.715,-2.916],[0.707106781,0,0,0.707106781],[0,0,0,0],[9E+09,9E+09,9E+09,9E+09,9E+09,9E+09]];
    CONST robtarget Target_Tap165_2690:=[[9.76,55.715,-20],[0.707106781,0,0,0.707106781],[0,0,0,0],[9E+09,9E+09,9E+09,9E+09,9E+09,9E+09]];
    CONST robtarget Target_Tap165_2700:=[[-2.908,55.576,-20],[0.707106781,0,0,0.707106781],[0,0,0,0],[9E+09,9E+09,9E+09,9E+09,9E+09,9E+09]];
    CONST robtarget Target_Tap165_2710:=[[-2.908,55.576,-3.031],[0.707106781,0,0,0.707106781],[0,0,0,0],[9E+09,9E+09,9E+09,9E+09,9E+09,9E+09]];
    CONST robtarget Target_Tap165_2720:=[[31.956,-5.382,-2.714],[0.707106781,0,0,0.707106781],[0,0,0,0],[9E+09,9E+09,9E+09,9E+09,9E+09,9E+09]];
    CONST robtarget Target_Tap165_2730:=[[34.985,-12.838,-2.687],[0.707106781,0,0,0.707106781],[0,0,0,0],[9E+09,9E+09,9E+09,9E+09,9E+09,9E+09]];
    CONST robtarget Target_Tap165_2740:=[[36.379,-19.375,-2.674],[0.707106781,0,0,0.707106781],[0,0,0,0],[9E+09,9E+09,9E+09,9E+09,9E+09,9E+09]];
    CONST robtarget Target_Tap165_2750:=[[36.379,-19.375,-19.674],[0.707106781,0,0,0.707106781],[0,0,0,0],[9E+09,9E+09,9E+09,9E+09,9E+09,9E+09]];
    CONST robtarget Target_Tap165_2760:=[[36.045,-22.924,-20],[0.707106781,0,0,0.707106781],[0,0,0,0],[9E+09,9E+09,9E+09,9E+09,9E+09,9E+09]];
    CONST robtarget Target_Tap165_2770:=[[36.045,-22.924,-2.677],[0.707106781,0,0,0.707106781],[0,0,0,0],[9E+09,9E+09,9E+09,9E+09,9E+09,9E+09]];
    CONST robtarget Target_Tap165_2780:=[[29.807,-37.797,-2.734],[0.707106781,0,0,0.707106781],[0,0,0,0],[9E+09,9E+09,9E+09,9E+09,9E+09,9E+09]];
    CONST robtarget Target_Tap165_2790:=[[16.78,-44.513,-2.852],[0.707106781,0,0,0.707106781],[0,0,0,0],[9E+09,9E+09,9E+09,9E+09,9E+09,9E+09]];
    CONST robtarget Target_Tap165_2800:=[[16.78,-44.513,-20],[0.707106781,0,0,0.707106781],[0,0,0,0],[9E+09,9E+09,9E+09,9E+09,9E+09,9E+09]];
    CONST robtarget Target_Tap165_2810:=[[13.526,-45.149,-20],[0.707106781,0,0,0.707106781],[0,0,0,0],[9E+09,9E+09,9E+09,9E+09,9E+09,9E+09]];
    CONST robtarget Target_Tap165_2820:=[[13.421,-44.964,-2.882],[0.707106781,0,0,0.707106781],[0,0,0,0],[9E+09,9E+09,9E+09,9E+09,9E+09,9E+09]];
    CONST robtarget Target_Tap165_2830:=[[1.129,-39.229,-2.994],[0.707106781,0,0,0.707106781],[0,0,0,0],[9E+09,9E+09,9E+09,9E+09,9E+09,9E+09]];
    CONST robtarget Target_Tap165_2840:=[[-6.679,-23.394,-3.065],[0.707106781,0,0,0.707106781],[0,0,0,0],[9E+09,9E+09,9E+09,9E+09,9E+09,9E+09]];
    CONST robtarget Target_Tap165_2850:=[[-6.679,-23.394,-20],[0.707106781,0,0,0.707106781],[0,0,0,0],[9E+09,9E+09,9E+09,9E+09,9E+09,9E+09]];
    CONST robtarget Target_Tap165_2860:=[[-5.981,-19.848,-20],[0.707106781,0,0,0.707106781],[0,0,0,0],[9E+09,9E+09,9E+09,9E+09,9E+09,9E+09]];
    CONST robtarget Target_Tap165_2870:=[[-5.981,-19.848,-3.058],[0.707106781,0,0,0.707106781],[0,0,0,0],[9E+09,9E+09,9E+09,9E+09,9E+09,9E+09]];
    CONST robtarget Target_Tap165_2880:=[[-0.37,-6.415,-3.007],[0.707106781,0,0,0.707106781],[0,0,0,0],[9E+09,9E+09,9E+09,9E+09,9E+09,9E+09]];
    CONST robtarget Target_Tap165_2890:=[[12.813,1.871,-2.888],[0.707106781,0,0,0.707106781],[0,0,0,0],[9E+09,9E+09,9E+09,9E+09,9E+09,9E+09]];
    CONST robtarget Target_Tap165_2900:=[[12.813,1.871,-20],[0.707106781,0,0,0.707106781],[0,0,0,0],[9E+09,9E+09,9E+09,9E+09,9E+09,9E+09]];
    CONST robtarget Target_Tap165_2910:=[[16.997,1.434,-20],[0.707106781,0,0,0.707106781],[0,0,0,0],[9E+09,9E+09,9E+09,9E+09,9E+09,9E+09]];
    CONST robtarget Target_Tap165_2920:=[[17.439,0.948,-2.846],[0.707106781,0,0,0.707106781],[0,0,0,0],[9E+09,9E+09,9E+09,9E+09,9E+09,9E+09]];
    CONST robtarget Target_Tap165_2930:=[[19.767,0.332,-2.825],[0.707106781,0,0,0.707106781],[0,0,0,0],[9E+09,9E+09,9E+09,9E+09,9E+09,9E+09]];
    CONST robtarget Target_Tap165_2940:=[[19.767,0.332,-20],[0.707106781,0,0,0.707106781],[0,0,0,0],[9E+09,9E+09,9E+09,9E+09,9E+09,9E+09]];
    CONST robtarget Target_Tap165_2950:=[[60.223,56.408,-20],[0.707106781,0,0,0.707106781],[0,0,0,0],[9E+09,9E+09,9E+09,9E+09,9E+09,9E+09]];
    CONST robtarget Target_Tap165_2960:=[[60.469,56.266,-2.455],[0.707106781,0,0,0.707106781],[0,0,0,0],[9E+09,9E+09,9E+09,9E+09,9E+09,9E+09]];
    CONST robtarget Target_Tap165_2970:=[[62.722,-59.754,-2.435],[0.707106781,0,0,0.707106781],[0,0,0,0],[9E+09,9E+09,9E+09,9E+09,9E+09,9E+09]];
    CONST robtarget Target_Tap165_2980:=[[62.722,-59.754,-20],[0.707106781,0,0,0.707106781],[0,0,0,0],[9E+09,9E+09,9E+09,9E+09,9E+09,9E+09]];
    CONST robtarget Target_Tap165_2990:=[[73.286,-59.666,-20],[0.707106781,0,0,0.707106781],[0,0,0,0],[9E+09,9E+09,9E+09,9E+09,9E+09,9E+09]];
    CONST robtarget Target_Tap165_3000:=[[73.286,-59.666,-2.339],[0.707106781,0,0,0.707106781],[0,0,0,0],[9E+09,9E+09,9E+09,9E+09,9E+09,9E+09]];
    CONST robtarget Target_Tap165_3010:=[[71.814,39.623,-2.352],[0.707106781,0,0,0.707106781],[0,0,0,0],[9E+09,9E+09,9E+09,9E+09,9E+09,9E+09]];
    CONST robtarget Target_Tap165_3020:=[[71.814,39.623,-20],[0.707106781,0,0,0.707106781],[0,0,0,0],[9E+09,9E+09,9E+09,9E+09,9E+09,9E+09]];
    CONST robtarget Target_Tap165_3030:=[[78.65,30.644,-20],[0.707106781,0,0,0.707106781],[0,0,0,0],[9E+09,9E+09,9E+09,9E+09,9E+09,9E+09]];
    CONST robtarget Target_Tap165_3040:=[[78.621,30.633,-1.291],[0.707106781,0,0,0.707106781],[0,0,0,0],[9E+09,9E+09,9E+09,9E+09,9E+09,9E+09]];
    CONST robtarget Target_Tap165_3050:=[[94.477,21.265,-1.147],[0.707106781,0,0,0.707106781],[0,0,0,0],[9E+09,9E+09,9E+09,9E+09,9E+09,9E+09]];
    CONST robtarget Target_Tap165_3060:=[[94.477,21.265,-20],[0.707106781,0,0,0.707106781],[0,0,0,0],[9E+09,9E+09,9E+09,9E+09,9E+09,9E+09]];
    CONST robtarget Target_Tap165_3070:=[[94.322,35.286,-20],[0.707106781,0,0,0.707106781],[0,0,0,0],[9E+09,9E+09,9E+09,9E+09,9E+09,9E+09]];
    CONST robtarget Target_Tap165_3080:=[[94.322,35.286,-1.148],[0.707106781,0,0,0.707106781],[0,0,0,0],[9E+09,9E+09,9E+09,9E+09,9E+09,9E+09]];
    CONST robtarget Target_Tap165_3090:=[[78.506,43.661,-1.292],[0.707106781,0,0,0.707106781],[0,0,0,0],[9E+09,9E+09,9E+09,9E+09,9E+09,9E+09]];
    CONST robtarget Target_Tap165_3100:=[[78.506,43.661,-20],[0.707106781,0,0,0.707106781],[0,0,0,0],[9E+09,9E+09,9E+09,9E+09,9E+09,9E+09]];
    CONST robtarget Target_Tap165_3110:=[[75.243,46.029,-20],[0.707106781,0,0,0.707106781],[0,0,0,0],[9E+09,9E+09,9E+09,9E+09,9E+09,9E+09]];
    CONST robtarget Target_Tap165_3120:=[[75.243,46.029,-1.321],[0.707106781,0,0,0.707106781],[0,0,0,0],[9E+09,9E+09,9E+09,9E+09,9E+09,9E+09]];
    CONST robtarget Target_Tap165_3130:=[[67.781,49.992,-1.389],[0.707106781,0,0,0.707106781],[0,0,0,0],[9E+09,9E+09,9E+09,9E+09,9E+09,9E+09]];
    CONST robtarget Target_Tap165_3140:=[[67.781,49.992,-20],[0.707106781,0,0,0.707106781],[0,0,0,0],[9E+09,9E+09,9E+09,9E+09,9E+09,9E+09]];
    CONST robtarget Target_Tap165_3150:=[[56.202,80.137,-20],[0.707106781,0,0,0.707106781],[0,0,0,0],[9E+09,9E+09,9E+09,9E+09,9E+09,9E+09]];
    CONST robtarget Target_Tap165_3160:=[[56.202,80.137,-2.494],[0.707106781,0,0,0.707106781],[0,0,0,0],[9E+09,9E+09,9E+09,9E+09,9E+09,9E+09]];
    CONST robtarget Target_Tap165_3170:=[[53.465,81.455,-2.519],[0.707106781,0,0,0.707106781],[0,0,0,0],[9E+09,9E+09,9E+09,9E+09,9E+09,9E+09]];
    CONST robtarget Target_Tap165_3180:=[[49.521,71.139,-2.555],[0.707106781,0,0,0.707106781],[0,0,0,0],[9E+09,9E+09,9E+09,9E+09,9E+09,9E+09]];
    CONST robtarget Target_Tap165_3190:=[[49.521,71.139,-20],[0.707106781,0,0,0.707106781],[0,0,0,0],[9E+09,9E+09,9E+09,9E+09,9E+09,9E+09]];
    CONST robtarget Target_Tap165_3200:=[[39.552,74.801,-20],[0.707106781,0,0,0.707106781],[0,0,0,0],[9E+09,9E+09,9E+09,9E+09,9E+09,9E+09]];
    CONST robtarget Target_Tap165_3210:=[[39.552,74.801,-2.645],[0.707106781,0,0,0.707106781],[0,0,0,0],[9E+09,9E+09,9E+09,9E+09,9E+09,9E+09]];
    CONST robtarget Target_Tap165_3220:=[[44.756,76.049,-2.598],[0.707106781,0,0,0.707106781],[0,0,0,0],[9E+09,9E+09,9E+09,9E+09,9E+09,9E+09]];
    CONST robtarget Target_Tap165_3230:=[[44.52,80.6,-2.6],[0.707106781,0,0,0.707106781],[0,0,0,0],[9E+09,9E+09,9E+09,9E+09,9E+09,9E+09]];
    CONST robtarget Target_Tap165_3240:=[[46.649,83.798,-2.581],[0.707106781,0,0,0.707106781],[0,0,0,0],[9E+09,9E+09,9E+09,9E+09,9E+09,9E+09]];
    CONST robtarget Target_Tap165_3250:=[[42.536,87.667,-2.618],[0.707106781,0,0,0.707106781],[0,0,0,0],[9E+09,9E+09,9E+09,9E+09,9E+09,9E+09]];
    CONST robtarget Target_Tap165_3260:=[[38.725,85.158,-2.653],[0.707106781,0,0,0.707106781],[0,0,0,0],[9E+09,9E+09,9E+09,9E+09,9E+09,9E+09]];
    CONST robtarget Target_Tap165_3270:=[[39.298,82.281,-2.647],[0.707106781,0,0,0.707106781],[0,0,0,0],[9E+09,9E+09,9E+09,9E+09,9E+09,9E+09]];
    CONST robtarget Target_Tap165_3280:=[[36.784,79.231,-2.67],[0.707106781,0,0,0.707106781],[0,0,0,0],[9E+09,9E+09,9E+09,9E+09,9E+09,9E+09]];
    CONST robtarget Target_Tap165_3290:=[[39.921,74.652,-2.642],[0.707106781,0,0,0.707106781],[0,0,0,0],[9E+09,9E+09,9E+09,9E+09,9E+09,9E+09]];
    CONST robtarget Target_Tap165_3300:=[[39.921,74.652,-20],[0.707106781,0,0,0.707106781],[0,0,0,0],[9E+09,9E+09,9E+09,9E+09,9E+09,9E+09]];
    CONST robtarget Target_Tap165_3310:=[[27.241,88.04,-19.757],[0.707106781,0,0,0.707106781],[0,0,0,0],[9E+09,9E+09,9E+09,9E+09,9E+09,9E+09]];
    CONST robtarget Target_Tap165_3320:=[[27.241,88.04,-2.757],[0.707106781,0,0,0.707106781],[0,0,0,0],[9E+09,9E+09,9E+09,9E+09,9E+09,9E+09]];
    CONST robtarget Target_Tap165_3330:=[[29.772,91.072,-2.734],[0.707106781,0,0,0.707106781],[0,0,0,0],[9E+09,9E+09,9E+09,9E+09,9E+09,9E+09]];
    CONST robtarget Target_Tap165_3340:=[[32.669,88.163,-2.708],[0.707106781,0,0,0.707106781],[0,0,0,0],[9E+09,9E+09,9E+09,9E+09,9E+09,9E+09]];
    CONST robtarget Target_Tap165_3350:=[[32.383,81.461,-2.71],[0.707106781,0,0,0.707106781],[0,0,0,0],[9E+09,9E+09,9E+09,9E+09,9E+09,9E+09]];
    CONST robtarget Target_Tap165_3360:=[[27.258,78.483,-2.757],[0.707106781,0,0,0.707106781],[0,0,0,0],[9E+09,9E+09,9E+09,9E+09,9E+09,9E+09]];
    CONST robtarget Target_Tap165_3370:=[[24.482,83.536,-2.782],[0.707106781,0,0,0.707106781],[0,0,0,0],[9E+09,9E+09,9E+09,9E+09,9E+09,9E+09]];
    CONST robtarget Target_Tap165_3380:=[[26.464,86.513,-2.764],[0.707106781,0,0,0.707106781],[0,0,0,0],[9E+09,9E+09,9E+09,9E+09,9E+09,9E+09]];
    CONST robtarget Target_Tap165_3390:=[[30.559,85.02,-2.727],[0.707106781,0,0,0.707106781],[0,0,0,0],[9E+09,9E+09,9E+09,9E+09,9E+09,9E+09]];
    CONST robtarget Target_Tap165_3400:=[[30.559,85.02,-20],[0.707106781,0,0,0.707106781],[0,0,0,0],[9E+09,9E+09,9E+09,9E+09,9E+09,9E+09]];
    CONST robtarget Target_Tap165_3410:=[[21.625,90.89,-20],[0.707106781,0,0,0.707106781],[0,0,0,0],[9E+09,9E+09,9E+09,9E+09,9E+09,9E+09]];
    CONST robtarget Target_Tap165_3420:=[[21.647,91.122,-2.808],[0.707106781,0,0,0.707106781],[0,0,0,0],[9E+09,9E+09,9E+09,9E+09,9E+09,9E+09]];
    CONST robtarget Target_Tap165_3430:=[[18.356,91.432,-2.838],[0.707106781,0,0,0.707106781],[0,0,0,0],[9E+09,9E+09,9E+09,9E+09,9E+09,9E+09]];
    CONST robtarget Target_Tap165_3440:=[[17.147,80.427,-2.848],[0.707106781,0,0,0.707106781],[0,0,0,0],[9E+09,9E+09,9E+09,9E+09,9E+09,9E+09]];
    CONST robtarget Target_Tap165_3450:=[[17.147,80.427,-20],[0.707106781,0,0,0.707106781],[0,0,0,0],[9E+09,9E+09,9E+09,9E+09,9E+09,9E+09]];
    CONST robtarget Target_Tap165_3460:=[[7.008,87.14,-20],[0.707106781,0,0,0.707106781],[0,0,0,0],[9E+09,9E+09,9E+09,9E+09,9E+09,9E+09]];
    CONST robtarget Target_Tap165_3470:=[[7.008,87.14,-2.941],[0.707106781,0,0,0.707106781],[0,0,0,0],[9E+09,9E+09,9E+09,9E+09,9E+09,9E+09]];
    CONST robtarget Target_Tap165_3480:=[[-0.038,87.612,-3.004],[0.707106781,0,0,0.707106781],[0,0,0,0],[9E+09,9E+09,9E+09,9E+09,9E+09,9E+09]];
    CONST robtarget Target_Tap165_3490:=[[-0.038,87.612,-20],[0.707106781,0,0,0.707106781],[0,0,0,0],[9E+09,9E+09,9E+09,9E+09,9E+09,9E+09]];
    CONST robtarget Target_Tap165_3500:=[[-11.27,89.538,-20],[0.707106781,0,0,0.707106781],[0,0,0,0],[9E+09,9E+09,9E+09,9E+09,9E+09,9E+09]];
    CONST robtarget Target_Tap165_3510:=[[-11.27,89.538,-3.106],[0.707106781,0,0,0.707106781],[0,0,0,0],[9E+09,9E+09,9E+09,9E+09,9E+09,9E+09]];
    CONST robtarget Target_Tap165_3520:=[[-15.219,93.483,-3.142],[0.707106781,0,0,0.707106781],[0,0,0,0],[9E+09,9E+09,9E+09,9E+09,9E+09,9E+09]];
    CONST robtarget Target_Tap165_3530:=[[-18.088,89.352,-3.168],[0.707106781,0,0,0.707106781],[0,0,0,0],[9E+09,9E+09,9E+09,9E+09,9E+09,9E+09]];
    CONST robtarget Target_Tap165_3540:=[[-9.511,81.207,-3.091],[0.707106781,0,0,0.707106781],[0,0,0,0],[9E+09,9E+09,9E+09,9E+09,9E+09,9E+09]];
    CONST robtarget Target_Tap165_3550:=[[-17.167,80.271,-3.16],[0.707106781,0,0,0.707106781],[0,0,0,0],[9E+09,9E+09,9E+09,9E+09,9E+09,9E+09]];
    CONST robtarget Target_Tap165_3560:=[[-17.167,80.271,-20],[0.707106781,0,0,0.707106781],[0,0,0,0],[9E+09,9E+09,9E+09,9E+09,9E+09,9E+09]];
    CONST robtarget Target_Tap165_3570:=[[-24.92,78.639,-20],[0.707106781,0,0,0.707106781],[0,0,0,0],[9E+09,9E+09,9E+09,9E+09,9E+09,9E+09]];
    CONST robtarget Target_Tap165_3580:=[[-24.92,78.639,-3.23],[0.707106781,0,0,0.707106781],[0,0,0,0],[9E+09,9E+09,9E+09,9E+09,9E+09,9E+09]];
    CONST robtarget Target_Tap165_3590:=[[-30.754,83.177,-3.283],[0.707106781,0,0,0.707106781],[0,0,0,0],[9E+09,9E+09,9E+09,9E+09,9E+09,9E+09]];
    CONST robtarget Target_Tap165_3600:=[[-27.506,91.364,-3.254],[0.707106781,0,0,0.707106781],[0,0,0,0],[9E+09,9E+09,9E+09,9E+09,9E+09,9E+09]];
    CONST robtarget Target_Tap165_3610:=[[-21.848,85.889,-3.202],[0.707106781,0,0,0.707106781],[0,0,0,0],[9E+09,9E+09,9E+09,9E+09,9E+09,9E+09]];
    CONST robtarget Target_Tap165_3620:=[[-24.92,78.639,-3.23],[0.707106781,0,0,0.707106781],[0,0,0,0],[9E+09,9E+09,9E+09,9E+09,9E+09,9E+09]];
    CONST robtarget Target_Tap165_3630:=[[-24.92,78.639,-20],[0.707106781,0,0,0.707106781],[0,0,0,0],[9E+09,9E+09,9E+09,9E+09,9E+09,9E+09]];
    CONST robtarget Target_Tap165_3640:=[[-36.608,84.296,-20],[0.707106781,0,0,0.707106781],[0,0,0,0],[9E+09,9E+09,9E+09,9E+09,9E+09,9E+09]];
    CONST robtarget Target_Tap165_3650:=[[-36.608,84.296,-3.336],[0.707106781,0,0,0.707106781],[0,0,0,0],[9E+09,9E+09,9E+09,9E+09,9E+09,9E+09]];
    CONST robtarget Target_Tap165_3660:=[[-40.159,87.789,-3.369],[0.707106781,0,0,0.707106781],[0,0,0,0],[9E+09,9E+09,9E+09,9E+09,9E+09,9E+09]];
    CONST robtarget Target_Tap165_3670:=[[-42.988,82.686,-3.394],[0.707106781,0,0,0.707106781],[0,0,0,0],[9E+09,9E+09,9E+09,9E+09,9E+09,9E+09]];
    CONST robtarget Target_Tap165_3680:=[[-33.051,76.713,-3.304],[0.707106781,0,0,0.707106781],[0,0,0,0],[9E+09,9E+09,9E+09,9E+09,9E+09,9E+09]];
    CONST robtarget Target_Tap165_3690:=[[-40.635,74.105,-3.373],[0.707106781,0,0,0.707106781],[0,0,0,0],[9E+09,9E+09,9E+09,9E+09,9E+09,9E+09]];
    CONST robtarget Target_Tap165_3700:=[[-40.661,74.141,-20],[0.707106781,0,0,0.707106781],[0,0,0,0],[9E+09,9E+09,9E+09,9E+09,9E+09,9E+09]];
    CONST robtarget Target_Tap165_3710:=[[-53.556,78.259,-20],[0.707106781,0,0,0.707106781],[0,0,0,0],[9E+09,9E+09,9E+09,9E+09,9E+09,9E+09]];
    CONST robtarget Target_Tap165_3720:=[[-53.519,78.274,-3.49],[0.707106781,0,0,0.707106781],[0,0,0,0],[9E+09,9E+09,9E+09,9E+09,9E+09,9E+09]];
    CONST robtarget Target_Tap165_3730:=[[-52.003,83.061,-3.476],[0.707106781,0,0,0.707106781],[0,0,0,0],[9E+09,9E+09,9E+09,9E+09,9E+09,9E+09]];
    CONST robtarget Target_Tap165_3740:=[[-47.618,81.007,-3.436],[0.707106781,0,0,0.707106781],[0,0,0,0],[9E+09,9E+09,9E+09,9E+09,9E+09,9E+09]];
    CONST robtarget Target_Tap165_3750:=[[-45.613,75.613,-3.418],[0.707106781,0,0,0.707106781],[0,0,0,0],[9E+09,9E+09,9E+09,9E+09,9E+09,9E+09]];
    CONST robtarget Target_Tap165_3760:=[[-48.776,70.343,-3.447],[0.707106781,0,0,0.707106781],[0,0,0,0],[9E+09,9E+09,9E+09,9E+09,9E+09,9E+09]];
    CONST robtarget Target_Tap165_3770:=[[-53.474,73.502,-3.489],[0.707106781,0,0,0.707106781],[0,0,0,0],[9E+09,9E+09,9E+09,9E+09,9E+09,9E+09]];
    CONST robtarget Target_Tap165_3780:=[[-52.696,77.199,-3.482],[0.707106781,0,0,0.707106781],[0,0,0,0],[9E+09,9E+09,9E+09,9E+09,9E+09,9E+09]];
    CONST robtarget Target_Tap165_3790:=[[-49.263,78.004,-3.451],[0.707106781,0,0,0.707106781],[0,0,0,0],[9E+09,9E+09,9E+09,9E+09,9E+09,9E+09]];
    CONST robtarget Target_Tap165_3800:=[[-49.263,78.004,-20],[0.707106781,0,0,0.707106781],[0,0,0,0],[9E+09,9E+09,9E+09,9E+09,9E+09,9E+09]];
    CONST robtarget p_contacto_165{319}:=[Target_Tap165_20, Target_Tap165_30, Target_Tap165_40, Target_Tap165_50, Target_Tap165_60, Target_Tap165_70,
                                       Target_Tap165_80, Target_Tap165_100, Target_Tap165_110, Target_Tap165_120, Target_Tap165_130, Target_Tap165_140,
                                       Target_Tap165_150, Target_Tap165_160, Target_Tap165_170, Target_Tap165_190, Target_Tap165_200, Target_Tap165_210,
                                       Target_Tap165_220, Target_Tap165_230, Target_Tap165_240, Target_Tap165_260, Target_Tap165_270, Target_Tap165_280,
                                       Target_Tap165_290, Target_Tap165_300, Target_Tap165_310, Target_Tap165_320, Target_Tap165_340, Target_Tap165_350,
                                       Target_Tap165_360, Target_Tap165_380, Target_Tap165_390, Target_Tap165_400, Target_Tap165_410, Target_Tap165_420,
                                       Target_Tap165_430, Target_Tap165_440, Target_Tap165_450, Target_Tap165_470, Target_Tap165_480, Target_Tap165_490,
                                       Target_Tap165_500, Target_Tap165_510, Target_Tap165_520, Target_Tap165_530, Target_Tap165_540, Target_Tap165_560,
                                       Target_Tap165_570, Target_Tap165_580, Target_Tap165_590, Target_Tap165_600, Target_Tap165_610, Target_Tap165_620,
                                       Target_Tap165_630, Target_Tap165_650, Target_Tap165_660, Target_Tap165_670, Target_Tap165_680, Target_Tap165_690,
                                       Target_Tap165_700, Target_Tap165_710, Target_Tap165_720, Target_Tap165_740, Target_Tap165_750, Target_Tap165_760,
                                       Target_Tap165_770, Target_Tap165_780, Target_Tap165_790, Target_Tap165_800, Target_Tap165_820, Target_Tap165_830,
                                       Target_Tap165_840, Target_Tap165_860, Target_Tap165_870, Target_Tap165_880, Target_Tap165_890, Target_Tap165_900,
                                       Target_Tap165_910, Target_Tap165_920, Target_Tap165_940, Target_Tap165_950, Target_Tap165_960, Target_Tap165_970,
                                       Target_Tap165_980, Target_Tap165_990, Target_Tap165_1000, Target_Tap165_1010, Target_Tap165_1020, Target_Tap165_1030,
                                       Target_Tap165_1050, Target_Tap165_1060, Target_Tap165_1070, Target_Tap165_1080, Target_Tap165_1090, Target_Tap165_1100,
                                       Target_Tap165_1110, Target_Tap165_1130, Target_Tap165_1140, Target_Tap165_1150, Target_Tap165_1160, Target_Tap165_1170,
                                       Target_Tap165_1180, Target_Tap165_1190, Target_Tap165_1210, Target_Tap165_1220, Target_Tap165_1230, Target_Tap165_1250,
                                       Target_Tap165_1260, Target_Tap165_1280, Target_Tap165_1290, Target_Tap165_1300, Target_Tap165_1310, Target_Tap165_1320,
                                       Target_Tap165_1330, Target_Tap165_1340, Target_Tap165_1360, Target_Tap165_1370, Target_Tap165_1380, Target_Tap165_1390,
                                       Target_Tap165_1400, Target_Tap165_1420, Target_Tap165_1430, Target_Tap165_1440, Target_Tap165_1460, Target_Tap165_1470,
                                       Target_Tap165_1480, Target_Tap165_1500, Target_Tap165_1510, Target_Tap165_1520, Target_Tap165_1530, Target_Tap165_1540,
                                       Target_Tap165_1550, Target_Tap165_1560, Target_Tap165_1570, Target_Tap165_1590, Target_Tap165_1600, Target_Tap165_1610,
                                       Target_Tap165_1620, Target_Tap165_1640, Target_Tap165_1650, Target_Tap165_1660, Target_Tap165_1670, Target_Tap165_1690,
                                       Target_Tap165_1700, Target_Tap165_1710, Target_Tap165_1720, Target_Tap165_1740, Target_Tap165_1750, Target_Tap165_1760,
                                       Target_Tap165_1780, Target_Tap165_1790, Target_Tap165_1800, Target_Tap165_1810, Target_Tap165_1830, Target_Tap165_1840,
                                       Target_Tap165_1850, Target_Tap165_1860, Target_Tap165_1880, Target_Tap165_1890, Target_Tap165_1900, Target_Tap165_1910,
                                       Target_Tap165_1930, Target_Tap165_1940, Target_Tap165_1950, Target_Tap165_1960, Target_Tap165_1970, Target_Tap165_1980,
                                       Target_Tap165_1990, Target_Tap165_2000, Target_Tap165_2020, Target_Tap165_2030, Target_Tap165_2040, Target_Tap165_2050,
                                       Target_Tap165_2060, Target_Tap165_2070, Target_Tap165_2080, Target_Tap165_2090, Target_Tap165_2110, Target_Tap165_2120,
                                       Target_Tap165_2130, Target_Tap165_2140, Target_Tap165_2150, Target_Tap165_2160, Target_Tap165_2180, Target_Tap165_2190,
                                       Target_Tap165_2200, Target_Tap165_2210, Target_Tap165_2220, Target_Tap165_2230, Target_Tap165_2250, Target_Tap165_2260,
                                       Target_Tap165_2270, Target_Tap165_2280, Target_Tap165_2290, Target_Tap165_2300, Target_Tap165_2310, Target_Tap165_2320,
                                       Target_Tap165_2340, Target_Tap165_2350, Target_Tap165_2360, Target_Tap165_2380, Target_Tap165_2390, Target_Tap165_2400,
                                       Target_Tap165_2420, Target_Tap165_2430, Target_Tap165_2440, Target_Tap165_2460, Target_Tap165_2470, Target_Tap165_2480,
                                       Target_Tap165_2500, Target_Tap165_2510, Target_Tap165_2520, Target_Tap165_2530, Target_Tap165_2550, Target_Tap165_2560,
                                       Target_Tap165_2570, Target_Tap165_2580, Target_Tap165_2600, Target_Tap165_2610, Target_Tap165_2620, Target_Tap165_2630,
                                       Target_Tap165_2650, Target_Tap165_2660, Target_Tap165_2670, Target_Tap165_2680, Target_Tap165_2690, Target_Tap165_2710,
                                       Target_Tap165_2720, Target_Tap165_2730, Target_Tap165_2740, Target_Tap165_2750, Target_Tap165_2770, Target_Tap165_2780,
                                       Target_Tap165_2790, Target_Tap165_2800, Target_Tap165_2820, Target_Tap165_2830, Target_Tap165_2840, Target_Tap165_2850,
                                       Target_Tap165_2870, Target_Tap165_2880, Target_Tap165_2890, Target_Tap165_2900, Target_Tap165_2920, Target_Tap165_2930,
                                       Target_Tap165_2940, Target_Tap165_2960, Target_Tap165_2970, Target_Tap165_2980, Target_Tap165_3000, Target_Tap165_3010,
                                       Target_Tap165_3020, Target_Tap165_3040, Target_Tap165_3050, Target_Tap165_3060, Target_Tap165_3080, Target_Tap165_3090,
                                       Target_Tap165_3100, Target_Tap165_3120, Target_Tap165_3130, Target_Tap165_3140, Target_Tap165_3160, Target_Tap165_3170,
                                       Target_Tap165_3180, Target_Tap165_3190, Target_Tap165_3210, Target_Tap165_3220, Target_Tap165_3230, Target_Tap165_3240,
                                       Target_Tap165_3250, Target_Tap165_3260, Target_Tap165_3270, Target_Tap165_3280, Target_Tap165_3290, Target_Tap165_3300,
                                       Target_Tap165_3320, Target_Tap165_3330, Target_Tap165_3340, Target_Tap165_3350, Target_Tap165_3360, Target_Tap165_3370,
                                       Target_Tap165_3380, Target_Tap165_3390, Target_Tap165_3400, Target_Tap165_3420, Target_Tap165_3430, Target_Tap165_3440,
                                       Target_Tap165_3450, Target_Tap165_3470, Target_Tap165_3480, Target_Tap165_3490, Target_Tap165_3510, Target_Tap165_3520,
                                       Target_Tap165_3530, Target_Tap165_3540, Target_Tap165_3550, Target_Tap165_3560, Target_Tap165_3580, Target_Tap165_3590,
                                       Target_Tap165_3600, Target_Tap165_3610, Target_Tap165_3620, Target_Tap165_3630, Target_Tap165_3650, Target_Tap165_3660,
                                       Target_Tap165_3670, Target_Tap165_3680, Target_Tap165_3690, Target_Tap165_3700, Target_Tap165_3720, Target_Tap165_3730,
                                       Target_Tap165_3740, Target_Tap165_3750, Target_Tap165_3760, Target_Tap165_3770, Target_Tap165_3780, Target_Tap165_3790,
                                       Target_Tap165_3800];
    CONST robtarget p_vacio_165{61}:=[Target_Tap165_10, Target_Tap165_90, Target_Tap165_180, Target_Tap165_250, Target_Tap165_330, Target_Tap165_370,
                                     Target_Tap165_460, Target_Tap165_550, Target_Tap165_640, Target_Tap165_730, Target_Tap165_810, Target_Tap165_850,
                                     Target_Tap165_930, Target_Tap165_1040, Target_Tap165_1120, Target_Tap165_1200, Target_Tap165_1240, Target_Tap165_1270,
                                     Target_Tap165_1350, Target_Tap165_1410, Target_Tap165_1450, Target_Tap165_1490, Target_Tap165_1580, Target_Tap165_1630,
                                     Target_Tap165_1680, Target_Tap165_1730, Target_Tap165_1770, Target_Tap165_1820, Target_Tap165_1870, Target_Tap165_1920,
                                     Target_Tap165_2010, Target_Tap165_2100, Target_Tap165_2170, Target_Tap165_2240, Target_Tap165_2330, Target_Tap165_2370,
                                     Target_Tap165_2410, Target_Tap165_2450, Target_Tap165_2490, Target_Tap165_2540, Target_Tap165_2590, Target_Tap165_2640,
                                     Target_Tap165_2700, Target_Tap165_2760, Target_Tap165_2810, Target_Tap165_2860, Target_Tap165_2910, Target_Tap165_2950,
                                     Target_Tap165_2990, Target_Tap165_3030, Target_Tap165_3070, Target_Tap165_3110, Target_Tap165_3150, Target_Tap165_3200,
                                     Target_Tap165_3310, Target_Tap165_3410, Target_Tap165_3460, Target_Tap165_3500, Target_Tap165_3570, Target_Tap165_3640,
                                     Target_Tap165_3710];

    PROC Decorar_Ing165(PERS wobjdata WO_Pastel)
        Mover_en_vacio;
        MoveJ Target_Home_10,Vel_Vacio_Rap,Z_Vacio_Rap,Prototipo_JSDaleman\WObj:=wobj0;
        ReiniciarIndices;
        path_contacto_actual:="p_contacto_165";
        path_vacio_actual:="p_vacio_165";
        Path_Tapa_165ing WO_Pastel;
        Mover_en_vacio;
        MoveJ Target_Home_10,Vel_Vacio_Rap,Z_Vacio_Rap,Prototipo_JSDaleman\WObj:=wobj0;
    ENDPROC
    PROC Path_Tapa_165ing(PERS wobjdata WO_Pastel)
        Path_vacio_ejecucion p_vacio_165, 1, WO_Pastel, FALSE;
        Path_contacto_ejecucion p_contacto_165, 1, 7, WO_Pastel, TRUE;
        Path_vacio_ejecucion p_vacio_165, 2, WO_Pastel, FALSE;
        index_vacio_destino:=15;
        Path_contacto_ejecucion p_contacto_165, 8, 10, WO_Pastel, FALSE;
        Mover_en_contacto;
        TriggC p_contacto_165{11},p_contacto_165{12},Vel_Proceso,triggContactoCir,Z_Proceso,Prototipo_JSDaleman\WObj:=WO_Pastel;
        TriggC p_contacto_165{13},p_contacto_165{14},Vel_Proceso,triggContactoCir,Z_Proceso,Prototipo_JSDaleman\WObj:=WO_Pastel;
        Mover_a_vacio;
        TriggL p_contacto_165{15},Vel_Acercamiento,triggContacto,Z_Acercamiento,Prototipo_JSDaleman\WObj:=WO_Pastel;
        Path_vacio_ejecucion p_vacio_165, 3, WO_Pastel, FALSE;
        index_vacio_destino:=21;
        Mover_a_contacto;
        TriggL p_contacto_165{16},Vel_Acercamiento,triggContacto,Z_Acercamiento,Prototipo_JSDaleman\WObj:=WO_Pastel;
        Mover_en_contacto;
        TriggC p_contacto_165{17},p_contacto_165{18},Vel_Proceso,triggContactoCir,Z_Proceso,Prototipo_JSDaleman\WObj:=WO_Pastel;
        TriggC p_contacto_165{19},p_contacto_165{20},Vel_Proceso,triggContactoCir,Z_Proceso,Prototipo_JSDaleman\WObj:=WO_Pastel;
        Mover_a_vacio;
        TriggL p_contacto_165{21},Vel_Acercamiento,triggContacto,Z_Acercamiento,Prototipo_JSDaleman\WObj:=WO_Pastel;
        Path_vacio_ejecucion p_vacio_165, 4, WO_Pastel, FALSE;
        index_vacio_destino:=28;
        Path_contacto_ejecucion p_contacto_165, 22, 23, WO_Pastel, FALSE;
        Mover_en_contacto;
        TriggC p_contacto_165{24},p_contacto_165{25},Vel_Proceso,triggContactoCir,Z_Proceso,Prototipo_JSDaleman\WObj:=WO_Pastel;
        TriggL p_contacto_165{26},Vel_Proceso,triggContacto,Z_Proceso,Prototipo_JSDaleman\WObj:=WO_Pastel;
        TriggL p_contacto_165{27},Vel_Proceso,triggContacto,Z_Proceso,Prototipo_JSDaleman\WObj:=WO_Pastel;
        Mover_a_vacio;
        TriggL p_contacto_165{28},Vel_Acercamiento,triggContacto,Z_Acercamiento,Prototipo_JSDaleman\WObj:=WO_Pastel;
        Path_vacio_ejecucion p_vacio_165, 5, WO_Pastel, FALSE;
        Path_contacto_ejecucion p_contacto_165, 29, 31, WO_Pastel, TRUE;
        Path_vacio_ejecucion p_vacio_165, 6, WO_Pastel, FALSE;
        Path_contacto_ejecucion p_contacto_165, 32, 39, WO_Pastel, TRUE;
        Path_vacio_ejecucion p_vacio_165, 7, WO_Pastel, FALSE;
        index_vacio_destino:=47;
        Path_contacto_ejecucion p_contacto_165, 40, 42, WO_Pastel, FALSE;
        Mover_en_contacto;
        TriggC p_contacto_165{43},p_contacto_165{44},Vel_Proceso,triggContactoCir,Z_Proceso,Prototipo_JSDaleman\WObj:=WO_Pastel;
        TriggC p_contacto_165{45},p_contacto_165{46},Vel_Proceso,triggContactoCir,Z_Proceso,Prototipo_JSDaleman\WObj:=WO_Pastel;
        Mover_a_vacio;
        TriggL p_contacto_165{47},Vel_Acercamiento,triggContacto,Z_Acercamiento,Prototipo_JSDaleman\WObj:=WO_Pastel;
        Path_vacio_ejecucion p_vacio_165, 8, WO_Pastel, FALSE;
        index_vacio_destino:=55;
        Path_contacto_ejecucion p_contacto_165, 48, 50, WO_Pastel, FALSE;
        Mover_en_contacto;
        TriggC p_contacto_165{51},p_contacto_165{52},Vel_Proceso,triggContactoCir,Z_Proceso,Prototipo_JSDaleman\WObj:=WO_Pastel;
        TriggC p_contacto_165{53},p_contacto_165{54},Vel_Proceso,triggContactoCir,Z_Proceso,Prototipo_JSDaleman\WObj:=WO_Pastel;
        Mover_a_vacio;
        TriggL p_contacto_165{55},Vel_Acercamiento,triggContacto,Z_Acercamiento,Prototipo_JSDaleman\WObj:=WO_Pastel;
        Path_vacio_ejecucion p_vacio_165, 9, WO_Pastel, FALSE;
        index_vacio_destino:=63;
        Path_contacto_ejecucion p_contacto_165, 56, 58, WO_Pastel, FALSE;
        Mover_en_contacto;
        TriggC p_contacto_165{59},p_contacto_165{60},Vel_Proceso,triggContactoCir,Z_Proceso,Prototipo_JSDaleman\WObj:=WO_Pastel;
        TriggC p_contacto_165{61},p_contacto_165{62},Vel_Proceso,triggContactoCir,Z_Proceso,Prototipo_JSDaleman\WObj:=WO_Pastel;
        Mover_a_vacio;
        TriggL p_contacto_165{63},Vel_Acercamiento,triggContacto,Z_Acercamiento,Prototipo_JSDaleman\WObj:=WO_Pastel;
        Path_vacio_ejecucion p_vacio_165, 10, WO_Pastel, FALSE;
        index_vacio_destino:=70;
        Mover_a_contacto;
        TriggL p_contacto_165{64},Vel_Acercamiento,triggContacto,Z_Acercamiento,Prototipo_JSDaleman\WObj:=WO_Pastel;
        Mover_en_contacto;
        TriggC p_contacto_165{65},p_contacto_165{66},Vel_Proceso,triggContactoCir,Z_Proceso,Prototipo_JSDaleman\WObj:=WO_Pastel;
        TriggC p_contacto_165{67},p_contacto_165{68},Vel_Proceso,triggContactoCir,Z_Proceso,Prototipo_JSDaleman\WObj:=WO_Pastel;
        TriggL p_contacto_165{69},Vel_Proceso,triggContacto,Z_Proceso,Prototipo_JSDaleman\WObj:=WO_Pastel;
        Mover_a_vacio;
        TriggL p_contacto_165{70},Vel_Acercamiento,triggContacto,Z_Acercamiento,Prototipo_JSDaleman\WObj:=WO_Pastel;
        Path_vacio_ejecucion p_vacio_165, 11, WO_Pastel, FALSE;
        Path_contacto_ejecucion p_contacto_165, 71, 73, WO_Pastel, TRUE;
        Path_vacio_ejecucion p_vacio_165, 12, WO_Pastel, FALSE;
        index_vacio_destino:=80;
        Path_contacto_ejecucion p_contacto_165, 74, 76, WO_Pastel, FALSE;
        Mover_en_contacto;
        TriggC p_contacto_165{77},p_contacto_165{78},Vel_Proceso,triggContactoCir,Z_Proceso,Prototipo_JSDaleman\WObj:=WO_Pastel;
        TriggL p_contacto_165{79},Vel_Proceso,triggContacto,Z_Proceso,Prototipo_JSDaleman\WObj:=WO_Pastel;
        Mover_a_vacio;
        TriggL p_contacto_165{80},Vel_Acercamiento,triggContacto,Z_Acercamiento,Prototipo_JSDaleman\WObj:=WO_Pastel;
        Path_vacio_ejecucion p_vacio_165, 13, WO_Pastel, FALSE;
        index_vacio_destino:=90;
        Mover_a_contacto;
        TriggL p_contacto_165{81},Vel_Acercamiento,triggContacto,Z_Acercamiento,Prototipo_JSDaleman\WObj:=WO_Pastel;
        Mover_en_contacto;
        TriggC p_contacto_165{82},p_contacto_165{83},Vel_Proceso,triggContactoCir,Z_Proceso,Prototipo_JSDaleman\WObj:=WO_Pastel;
        TriggL p_contacto_165{84},Vel_Proceso,triggContacto,Z_Proceso,Prototipo_JSDaleman\WObj:=WO_Pastel;
        TriggL p_contacto_165{85},Vel_Proceso,triggContacto,Z_Proceso,Prototipo_JSDaleman\WObj:=WO_Pastel;
        TriggC p_contacto_165{86},p_contacto_165{87},Vel_Proceso,triggContactoCir,Z_Proceso,Prototipo_JSDaleman\WObj:=WO_Pastel;
        TriggC p_contacto_165{88},p_contacto_165{89},Vel_Proceso,triggContactoCir,Z_Proceso,Prototipo_JSDaleman\WObj:=WO_Pastel;
        Mover_a_vacio;
        TriggL p_contacto_165{90},Vel_Acercamiento,triggContacto,Z_Acercamiento,Prototipo_JSDaleman\WObj:=WO_Pastel;
        Path_vacio_ejecucion p_vacio_165, 14, WO_Pastel, FALSE;
        index_vacio_destino:=97;
        Mover_a_contacto;
        TriggL p_contacto_165{91},Vel_Acercamiento,triggContacto,Z_Acercamiento,Prototipo_JSDaleman\WObj:=WO_Pastel;
        Mover_en_contacto;
        TriggC p_contacto_165{92},p_contacto_165{93},Vel_Proceso,triggContactoCir,Z_Proceso,Prototipo_JSDaleman\WObj:=WO_Pastel;
        TriggC p_contacto_165{94},p_contacto_165{95},Vel_Proceso,triggContactoCir,Z_Proceso,Prototipo_JSDaleman\WObj:=WO_Pastel;
        TriggL p_contacto_165{96},Vel_Proceso,triggContacto,Z_Proceso,Prototipo_JSDaleman\WObj:=WO_Pastel;
        Mover_a_vacio;
        TriggL p_contacto_165{97},Vel_Acercamiento,triggContacto,Z_Acercamiento,Prototipo_JSDaleman\WObj:=WO_Pastel;
        Path_vacio_ejecucion p_vacio_165, 15, WO_Pastel, FALSE;
        index_vacio_destino:=104;
        Path_contacto_ejecucion p_contacto_165, 98, 100, WO_Pastel, FALSE;
        Mover_en_contacto;
        TriggC p_contacto_165{101},p_contacto_165{102},Vel_Proceso,triggContactoCir,Z_Proceso,Prototipo_JSDaleman\WObj:=WO_Pastel;
        TriggL p_contacto_165{103},Vel_Proceso,triggContacto,Z_Proceso,Prototipo_JSDaleman\WObj:=WO_Pastel;
        Mover_a_vacio;
        TriggL p_contacto_165{104},Vel_Acercamiento,triggContacto,Z_Acercamiento,Prototipo_JSDaleman\WObj:=WO_Pastel;
        Path_vacio_ejecucion p_vacio_165, 16, WO_Pastel, FALSE;
        Path_contacto_ejecucion p_contacto_165, 105, 107, WO_Pastel, TRUE;
        Path_vacio_ejecucion p_vacio_165, 17, WO_Pastel, FALSE;
        Path_contacto_ejecucion p_contacto_165, 108, 109, WO_Pastel, TRUE;
        Path_vacio_ejecucion p_vacio_165, 18, WO_Pastel, FALSE;
        index_vacio_destino:=116;
        Mover_a_contacto;
        TriggL p_contacto_165{110},Vel_Acercamiento,triggContacto,Z_Acercamiento,Prototipo_JSDaleman\WObj:=WO_Pastel;
        Mover_en_contacto;
        TriggC p_contacto_165{111},p_contacto_165{112},Vel_Proceso,triggContactoCir,Z_Proceso,Prototipo_JSDaleman\WObj:=WO_Pastel;
        TriggC p_contacto_165{113},p_contacto_165{114},Vel_Proceso,triggContactoCir,Z_Proceso,Prototipo_JSDaleman\WObj:=WO_Pastel;
        TriggL p_contacto_165{115},Vel_Proceso,triggContacto,Z_Proceso,Prototipo_JSDaleman\WObj:=WO_Pastel;
        Mover_a_vacio;
        TriggL p_contacto_165{116},Vel_Acercamiento,triggContacto,Z_Acercamiento,Prototipo_JSDaleman\WObj:=WO_Pastel;
        Path_vacio_ejecucion p_vacio_165, 19, WO_Pastel, FALSE;
        Path_contacto_ejecucion p_contacto_165, 117, 121, WO_Pastel, TRUE;
        Path_vacio_ejecucion p_vacio_165, 20, WO_Pastel, FALSE;
        Path_contacto_ejecucion p_contacto_165, 122, 124, WO_Pastel, TRUE;
        Path_vacio_ejecucion p_vacio_165, 21, WO_Pastel, FALSE;
        Path_contacto_ejecucion p_contacto_165, 125, 127, WO_Pastel, TRUE;
        Path_vacio_ejecucion p_vacio_165, 22, WO_Pastel, FALSE;
        index_vacio_destino:=135;
        Path_contacto_ejecucion p_contacto_165, 128, 130, WO_Pastel, FALSE;
        Mover_en_contacto;
        TriggC p_contacto_165{131},p_contacto_165{132},Vel_Proceso,triggContactoCir,Z_Proceso,Prototipo_JSDaleman\WObj:=WO_Pastel;
        TriggC p_contacto_165{133},p_contacto_165{134},Vel_Proceso,triggContactoCir,Z_Proceso,Prototipo_JSDaleman\WObj:=WO_Pastel;
        Mover_a_vacio;
        TriggL p_contacto_165{135},Vel_Acercamiento,triggContacto,Z_Acercamiento,Prototipo_JSDaleman\WObj:=WO_Pastel;
        Path_vacio_ejecucion p_vacio_165, 23, WO_Pastel, FALSE;
        index_vacio_destino:=139;
        Mover_a_contacto;
        TriggL p_contacto_165{136},Vel_Acercamiento,triggContacto,Z_Acercamiento,Prototipo_JSDaleman\WObj:=WO_Pastel;
        Mover_en_contacto;
        TriggC p_contacto_165{137},p_contacto_165{138},Vel_Proceso,triggContactoCir,Z_Proceso,Prototipo_JSDaleman\WObj:=WO_Pastel;
        Mover_a_vacio;
        TriggL p_contacto_165{139},Vel_Acercamiento,triggContacto,Z_Acercamiento,Prototipo_JSDaleman\WObj:=WO_Pastel;
        Path_vacio_ejecucion p_vacio_165, 24, WO_Pastel, FALSE;
        index_vacio_destino:=143;
        Mover_a_contacto;
        TriggL p_contacto_165{140},Vel_Acercamiento,triggContacto,Z_Acercamiento,Prototipo_JSDaleman\WObj:=WO_Pastel;
        Mover_en_contacto;
        TriggC p_contacto_165{141},p_contacto_165{142},Vel_Proceso,triggContactoCir,Z_Proceso,Prototipo_JSDaleman\WObj:=WO_Pastel;
        Mover_a_vacio;
        TriggL p_contacto_165{143},Vel_Acercamiento,triggContacto,Z_Acercamiento,Prototipo_JSDaleman\WObj:=WO_Pastel;
        Path_vacio_ejecucion p_vacio_165, 25, WO_Pastel, FALSE;
        index_vacio_destino:=147;
        Mover_a_contacto;
        TriggL p_contacto_165{144},Vel_Acercamiento,triggContacto,Z_Acercamiento,Prototipo_JSDaleman\WObj:=WO_Pastel;
        Mover_en_contacto;
        TriggC p_contacto_165{145},p_contacto_165{146},Vel_Proceso,triggContactoCir,Z_Proceso,Prototipo_JSDaleman\WObj:=WO_Pastel;
        Mover_a_vacio;
        TriggL p_contacto_165{147},Vel_Acercamiento,triggContacto,Z_Acercamiento,Prototipo_JSDaleman\WObj:=WO_Pastel;
        Path_vacio_ejecucion p_vacio_165, 26, WO_Pastel, FALSE;
        Path_contacto_ejecucion p_contacto_165, 148, 150, WO_Pastel, TRUE;
        Path_vacio_ejecucion p_vacio_165, 27, WO_Pastel, FALSE;
        index_vacio_destino:=154;
        Mover_a_contacto;
        TriggL p_contacto_165{151},Vel_Acercamiento,triggContacto,Z_Acercamiento,Prototipo_JSDaleman\WObj:=WO_Pastel;
        Mover_en_contacto;
        TriggC p_contacto_165{152},p_contacto_165{153},Vel_Proceso,triggContactoCir,Z_Proceso,Prototipo_JSDaleman\WObj:=WO_Pastel;
        Mover_a_vacio;
        TriggL p_contacto_165{154},Vel_Acercamiento,triggContacto,Z_Acercamiento,Prototipo_JSDaleman\WObj:=WO_Pastel;
        Path_vacio_ejecucion p_vacio_165, 28, WO_Pastel, FALSE;
        index_vacio_destino:=158;
        Mover_a_contacto;
        TriggL p_contacto_165{155},Vel_Acercamiento,triggContacto,Z_Acercamiento,Prototipo_JSDaleman\WObj:=WO_Pastel;
        Mover_en_contacto;
        TriggC p_contacto_165{156},p_contacto_165{157},Vel_Proceso,triggContactoCir,Z_Proceso,Prototipo_JSDaleman\WObj:=WO_Pastel;
        Mover_a_vacio;
        TriggL p_contacto_165{158},Vel_Acercamiento,triggContacto,Z_Acercamiento,Prototipo_JSDaleman\WObj:=WO_Pastel;
        Path_vacio_ejecucion p_vacio_165, 29, WO_Pastel, FALSE;
        index_vacio_destino:=162;
        Mover_a_contacto;
        TriggL p_contacto_165{159},Vel_Acercamiento,triggContacto,Z_Acercamiento,Prototipo_JSDaleman\WObj:=WO_Pastel;
        Mover_en_contacto;
        TriggC p_contacto_165{160},p_contacto_165{161},Vel_Proceso,triggContactoCir,Z_Proceso,Prototipo_JSDaleman\WObj:=WO_Pastel;
        Mover_a_vacio;
        TriggL p_contacto_165{162},Vel_Acercamiento,triggContacto,Z_Acercamiento,Prototipo_JSDaleman\WObj:=WO_Pastel;
        Path_vacio_ejecucion p_vacio_165, 30, WO_Pastel, FALSE;
        index_vacio_destino:=170;
        Path_contacto_ejecucion p_contacto_165, 163, 165, WO_Pastel, FALSE;
        Mover_en_contacto;
        TriggC p_contacto_165{166},p_contacto_165{167},Vel_Proceso,triggContactoCir,Z_Proceso,Prototipo_JSDaleman\WObj:=WO_Pastel;
        TriggC p_contacto_165{168},p_contacto_165{169},Vel_Proceso,triggContactoCir,Z_Proceso,Prototipo_JSDaleman\WObj:=WO_Pastel;
        Mover_a_vacio;
        TriggL p_contacto_165{170},Vel_Acercamiento,triggContacto,Z_Acercamiento,Prototipo_JSDaleman\WObj:=WO_Pastel;
        Path_vacio_ejecucion p_vacio_165, 31, WO_Pastel, FALSE;
        index_vacio_destino:=178;
        Path_contacto_ejecucion p_contacto_165, 171, 173, WO_Pastel, FALSE;
        Mover_en_contacto;
        TriggC p_contacto_165{174},p_contacto_165{175},Vel_Proceso,triggContactoCir,Z_Proceso,Prototipo_JSDaleman\WObj:=WO_Pastel;
        TriggL p_contacto_165{176},Vel_Proceso,triggContacto,Z_Proceso,Prototipo_JSDaleman\WObj:=WO_Pastel;
        TriggL p_contacto_165{177},Vel_Proceso,triggContacto,Z_Proceso,Prototipo_JSDaleman\WObj:=WO_Pastel;
        Mover_a_vacio;
        TriggL p_contacto_165{178},Vel_Acercamiento,triggContacto,Z_Acercamiento,Prototipo_JSDaleman\WObj:=WO_Pastel;
        Path_vacio_ejecucion p_vacio_165, 32, WO_Pastel, FALSE;
        index_vacio_destino:=184;
        Mover_a_contacto;
        TriggL p_contacto_165{179},Vel_Acercamiento,triggContacto,Z_Acercamiento,Prototipo_JSDaleman\WObj:=WO_Pastel;
        Mover_en_contacto;
        TriggC p_contacto_165{180},p_contacto_165{181},Vel_Proceso,triggContactoCir,Z_Proceso,Prototipo_JSDaleman\WObj:=WO_Pastel;
        TriggC p_contacto_165{182},p_contacto_165{183},Vel_Proceso,triggContactoCir,Z_Proceso,Prototipo_JSDaleman\WObj:=WO_Pastel;
        Mover_a_vacio;
        TriggL p_contacto_165{184},Vel_Acercamiento,triggContacto,Z_Acercamiento,Prototipo_JSDaleman\WObj:=WO_Pastel;
        Path_vacio_ejecucion p_vacio_165, 33, WO_Pastel, FALSE;
        index_vacio_destino:=190;
        Mover_a_contacto;
        TriggL p_contacto_165{185},Vel_Acercamiento,triggContacto,Z_Acercamiento,Prototipo_JSDaleman\WObj:=WO_Pastel;
        Mover_en_contacto;
        TriggC p_contacto_165{186},p_contacto_165{187},Vel_Proceso,triggContactoCir,Z_Proceso,Prototipo_JSDaleman\WObj:=WO_Pastel;
        TriggC p_contacto_165{188},p_contacto_165{189},Vel_Proceso,triggContactoCir,Z_Proceso,Prototipo_JSDaleman\WObj:=WO_Pastel;
        Mover_a_vacio;
        TriggL p_contacto_165{190},Vel_Acercamiento,triggContacto,Z_Acercamiento,Prototipo_JSDaleman\WObj:=WO_Pastel;
        Path_vacio_ejecucion p_vacio_165, 34, WO_Pastel, FALSE;
        index_vacio_destino:=198;
        Mover_a_contacto;
        TriggL p_contacto_165{191},Vel_Acercamiento,triggContacto,Z_Acercamiento,Prototipo_JSDaleman\WObj:=WO_Pastel;
        Mover_en_contacto;
        TriggC p_contacto_165{192},p_contacto_165{193},Vel_Proceso,triggContactoCir,Z_Proceso,Prototipo_JSDaleman\WObj:=WO_Pastel;
        TriggL p_contacto_165{194},Vel_Proceso,triggContacto,Z_Proceso,Prototipo_JSDaleman\WObj:=WO_Pastel;
        TriggL p_contacto_165{195},Vel_Proceso,triggContacto,Z_Proceso,Prototipo_JSDaleman\WObj:=WO_Pastel;
        TriggC p_contacto_165{196},p_contacto_165{197},Vel_Proceso,triggContactoCir,Z_Proceso,Prototipo_JSDaleman\WObj:=WO_Pastel;
        Mover_a_vacio;
        TriggL p_contacto_165{198},Vel_Acercamiento,triggContacto,Z_Acercamiento,Prototipo_JSDaleman\WObj:=WO_Pastel;
        Path_vacio_ejecucion p_vacio_165, 35, WO_Pastel, FALSE;
        Path_contacto_ejecucion p_contacto_165, 199, 201, WO_Pastel, TRUE;
        Path_vacio_ejecucion p_vacio_165, 36, WO_Pastel, FALSE;
        Path_contacto_ejecucion p_contacto_165, 202, 204, WO_Pastel, TRUE;
        Path_vacio_ejecucion p_vacio_165, 37, WO_Pastel, FALSE;
        Path_contacto_ejecucion p_contacto_165, 205, 207, WO_Pastel, TRUE;
        Path_vacio_ejecucion p_vacio_165, 38, WO_Pastel, FALSE;
        Path_contacto_ejecucion p_contacto_165, 208, 210, WO_Pastel, TRUE;
        Path_vacio_ejecucion p_vacio_165, 39, WO_Pastel, FALSE;
        index_vacio_destino:=214;
        Mover_a_contacto;
        TriggL p_contacto_165{211},Vel_Acercamiento,triggContacto,Z_Acercamiento,Prototipo_JSDaleman\WObj:=WO_Pastel;
        Mover_en_contacto;
        TriggC p_contacto_165{212},p_contacto_165{213},Vel_Proceso,triggContactoCir,Z_Proceso,Prototipo_JSDaleman\WObj:=WO_Pastel;
        Mover_a_vacio;
        TriggL p_contacto_165{214},Vel_Acercamiento,triggContacto,Z_Acercamiento,Prototipo_JSDaleman\WObj:=WO_Pastel;
        Path_vacio_ejecucion p_vacio_165, 40, WO_Pastel, FALSE;
        index_vacio_destino:=218;
        Mover_a_contacto;
        TriggL p_contacto_165{215},Vel_Acercamiento,triggContacto,Z_Acercamiento,Prototipo_JSDaleman\WObj:=WO_Pastel;
        Mover_en_contacto;
        TriggC p_contacto_165{216},p_contacto_165{217},Vel_Proceso,triggContactoCir,Z_Proceso,Prototipo_JSDaleman\WObj:=WO_Pastel;
        Mover_a_vacio;
        TriggL p_contacto_165{218},Vel_Acercamiento,triggContacto,Z_Acercamiento,Prototipo_JSDaleman\WObj:=WO_Pastel;
        Path_vacio_ejecucion p_vacio_165, 41, WO_Pastel, FALSE;
        index_vacio_destino:=222;
        Mover_a_contacto;
        TriggL p_contacto_165{219},Vel_Acercamiento,triggContacto,Z_Acercamiento,Prototipo_JSDaleman\WObj:=WO_Pastel;
        Mover_en_contacto;
        TriggC p_contacto_165{220},p_contacto_165{221},Vel_Proceso,triggContactoCir,Z_Proceso,Prototipo_JSDaleman\WObj:=WO_Pastel;
        Mover_a_vacio;
        TriggL p_contacto_165{222},Vel_Acercamiento,triggContacto,Z_Acercamiento,Prototipo_JSDaleman\WObj:=WO_Pastel;
        Path_vacio_ejecucion p_vacio_165, 42, WO_Pastel, FALSE;
        index_vacio_destino:=227;
        Mover_a_contacto;
        TriggL p_contacto_165{223},Vel_Acercamiento,triggContacto,Z_Acercamiento,Prototipo_JSDaleman\WObj:=WO_Pastel;
        Mover_en_contacto;
        TriggC p_contacto_165{224},p_contacto_165{225},Vel_Proceso,triggContactoCir,Z_Proceso,Prototipo_JSDaleman\WObj:=WO_Pastel;
        TriggL p_contacto_165{226},Vel_Proceso,triggContacto,Z_Proceso,Prototipo_JSDaleman\WObj:=WO_Pastel;
        Mover_a_vacio;
        TriggL p_contacto_165{227},Vel_Acercamiento,triggContacto,Z_Acercamiento,Prototipo_JSDaleman\WObj:=WO_Pastel;
        Path_vacio_ejecucion p_vacio_165, 43, WO_Pastel, FALSE;
        index_vacio_destino:=232;
        Mover_a_contacto;
        TriggL p_contacto_165{228},Vel_Acercamiento,triggContacto,Z_Acercamiento,Prototipo_JSDaleman\WObj:=WO_Pastel;
        TriggL p_contacto_165{229},Vel_Proceso,triggContacto,Z_Proceso,Prototipo_JSDaleman\WObj:=WO_Pastel;
        TriggC p_contacto_165{230},p_contacto_165{231},Vel_Proceso,triggContactoCir,Z_Proceso,Prototipo_JSDaleman\WObj:=WO_Pastel;
        Mover_a_vacio;
        TriggL p_contacto_165{232},Vel_Acercamiento,triggContacto,Z_Acercamiento,Prototipo_JSDaleman\WObj:=WO_Pastel;
        Path_vacio_ejecucion p_vacio_165, 44, WO_Pastel, FALSE;
        index_vacio_destino:=236;
        Mover_a_contacto;
        TriggL p_contacto_165{233},Vel_Acercamiento,triggContacto,Z_Acercamiento,Prototipo_JSDaleman\WObj:=WO_Pastel;
        Mover_en_contacto;
        TriggC p_contacto_165{234},p_contacto_165{235},Vel_Proceso,triggContactoCir,Z_Proceso,Prototipo_JSDaleman\WObj:=WO_Pastel;
        Mover_a_vacio;
        TriggL p_contacto_165{236},Vel_Acercamiento,triggContacto,Z_Acercamiento,Prototipo_JSDaleman\WObj:=WO_Pastel;
        Path_vacio_ejecucion p_vacio_165, 45, WO_Pastel, FALSE;
        index_vacio_destino:=240;
        Mover_a_contacto;
        TriggL p_contacto_165{237},Vel_Acercamiento,triggContacto,Z_Acercamiento,Prototipo_JSDaleman\WObj:=WO_Pastel;
        Mover_en_contacto;
        TriggC p_contacto_165{238},p_contacto_165{239},Vel_Proceso,triggContactoCir,Z_Proceso,Prototipo_JSDaleman\WObj:=WO_Pastel;
        Mover_a_vacio;
        TriggL p_contacto_165{240},Vel_Acercamiento,triggContacto,Z_Acercamiento,Prototipo_JSDaleman\WObj:=WO_Pastel;
        Path_vacio_ejecucion p_vacio_165, 46, WO_Pastel, FALSE;
        index_vacio_destino:=244;
        Mover_a_contacto;
        TriggL p_contacto_165{241},Vel_Acercamiento,triggContacto,Z_Acercamiento,Prototipo_JSDaleman\WObj:=WO_Pastel;
        Mover_en_contacto;
        TriggC p_contacto_165{242},p_contacto_165{243},Vel_Proceso,triggContactoCir,Z_Proceso,Prototipo_JSDaleman\WObj:=WO_Pastel;
        Mover_a_vacio;
        TriggL p_contacto_165{244},Vel_Acercamiento,triggContacto,Z_Acercamiento,Prototipo_JSDaleman\WObj:=WO_Pastel;
        Path_vacio_ejecucion p_vacio_165, 47, WO_Pastel, FALSE;
        index_vacio_destino:=247;
        Mover_a_contacto;
        TriggL p_contacto_165{245},Vel_Acercamiento,triggContacto,Z_Acercamiento,Prototipo_JSDaleman\WObj:=WO_Pastel;
        Mover_en_contacto;
        TriggL p_contacto_165{246},Vel_Proceso,triggContacto,Z_Proceso,Prototipo_JSDaleman\WObj:=WO_Pastel;
        Mover_a_vacio;
        TriggL p_contacto_165{247},Vel_Acercamiento,triggContacto,Z_Acercamiento,Prototipo_JSDaleman\WObj:=WO_Pastel;
        Path_vacio_ejecucion p_vacio_165, 48, WO_Pastel, FALSE;
        Path_contacto_ejecucion p_contacto_165, 248, 250, WO_Pastel, TRUE;
        Path_vacio_ejecucion p_vacio_165, 49, WO_Pastel, FALSE;
        Path_contacto_ejecucion p_contacto_165, 251, 253, WO_Pastel, TRUE;
        Path_vacio_ejecucion p_vacio_165, 50, WO_Pastel, FALSE;
        Path_contacto_ejecucion p_contacto_165, 254, 256, WO_Pastel, TRUE;
        Path_vacio_ejecucion p_vacio_165, 51, WO_Pastel, FALSE;
        Path_contacto_ejecucion p_contacto_165, 257, 259, WO_Pastel, TRUE;
        Path_vacio_ejecucion p_vacio_165, 52, WO_Pastel, FALSE;
        Path_contacto_ejecucion p_contacto_165, 260, 262, WO_Pastel, TRUE;
        Path_vacio_ejecucion p_vacio_165, 53, WO_Pastel, FALSE;
        Path_contacto_ejecucion p_contacto_165, 263, 266, WO_Pastel, TRUE;
        Path_vacio_ejecucion p_vacio_165, 54, WO_Pastel, FALSE;
        index_vacio_destino:=276;
        Mover_a_contacto;
        TriggL p_contacto_165{267},Vel_Acercamiento,triggContacto,Z_Acercamiento,Prototipo_JSDaleman\WObj:=WO_Pastel;
        Mover_en_contacto;
        TriggC p_contacto_165{268},p_contacto_165{269},Vel_Proceso,triggContactoCir,Z_Proceso,Prototipo_JSDaleman\WObj:=WO_Pastel;
        TriggC p_contacto_165{270},p_contacto_165{271},Vel_Proceso,triggContactoCir,Z_Proceso,Prototipo_JSDaleman\WObj:=WO_Pastel;
        TriggC p_contacto_165{272},p_contacto_165{273},Vel_Proceso,triggContactoCir,Z_Proceso,Prototipo_JSDaleman\WObj:=WO_Pastel;
        TriggC p_contacto_165{274},p_contacto_165{275},Vel_Proceso,triggContactoCir,Z_Proceso,Prototipo_JSDaleman\WObj:=WO_Pastel;
        Mover_a_vacio;
        TriggL p_contacto_165{276},Vel_Acercamiento,triggContacto,Z_Acercamiento,Prototipo_JSDaleman\WObj:=WO_Pastel;
        Path_vacio_ejecucion p_vacio_165, 55, WO_Pastel, FALSE;
        index_vacio_destino:=285;
        Mover_a_contacto;
        TriggL p_contacto_165{277},Vel_Acercamiento,triggContacto,Z_Acercamiento,Prototipo_JSDaleman\WObj:=WO_Pastel;
        Mover_en_contacto;
        TriggC p_contacto_165{278},p_contacto_165{279},Vel_Proceso,triggContactoCir,Z_Proceso,Prototipo_JSDaleman\WObj:=WO_Pastel;
        TriggL p_contacto_165{280},Vel_Proceso,triggContacto,Z_Proceso,Prototipo_JSDaleman\WObj:=WO_Pastel;
        TriggC p_contacto_165{281},p_contacto_165{282},Vel_Proceso,triggContactoCir,Z_Proceso,Prototipo_JSDaleman\WObj:=WO_Pastel;
        TriggC p_contacto_165{283},p_contacto_165{284},Vel_Proceso,triggContactoCir,Z_Proceso,Prototipo_JSDaleman\WObj:=WO_Pastel;
        Mover_a_vacio;
        TriggL p_contacto_165{285},Vel_Acercamiento,triggContacto,Z_Acercamiento,Prototipo_JSDaleman\WObj:=WO_Pastel;
        Path_vacio_ejecucion p_vacio_165, 56, WO_Pastel, FALSE;
        Path_contacto_ejecucion p_contacto_165, 286, 289, WO_Pastel, TRUE;
        Path_vacio_ejecucion p_vacio_165, 57, WO_Pastel, FALSE;
        Path_contacto_ejecucion p_contacto_165, 290, 292, WO_Pastel, TRUE;
        Path_vacio_ejecucion p_vacio_165, 58, WO_Pastel, FALSE;
        index_vacio_destino:=298;
        Mover_a_contacto;
        TriggL p_contacto_165{293},Vel_Acercamiento,triggContacto,Z_Acercamiento,Prototipo_JSDaleman\WObj:=WO_Pastel;
        Mover_en_contacto;
        TriggC p_contacto_165{294},p_contacto_165{295},Vel_Proceso,triggContactoCir,Z_Proceso,Prototipo_JSDaleman\WObj:=WO_Pastel;
        TriggL p_contacto_165{296},Vel_Proceso,triggContacto,Z_Proceso,Prototipo_JSDaleman\WObj:=WO_Pastel;
        TriggL p_contacto_165{297},Vel_Proceso,triggContacto,Z_Proceso,Prototipo_JSDaleman\WObj:=WO_Pastel;
        Mover_a_vacio;
        TriggL p_contacto_165{298},Vel_Acercamiento,triggContacto,Z_Acercamiento,Prototipo_JSDaleman\WObj:=WO_Pastel;
        Path_vacio_ejecucion p_vacio_165, 59, WO_Pastel, FALSE;
        index_vacio_destino:=304;
        Mover_a_contacto;
        TriggL p_contacto_165{299},Vel_Acercamiento,triggContacto,Z_Acercamiento,Prototipo_JSDaleman\WObj:=WO_Pastel;
        Mover_en_contacto;
        TriggC p_contacto_165{300},p_contacto_165{301},Vel_Proceso,triggContactoCir,Z_Proceso,Prototipo_JSDaleman\WObj:=WO_Pastel;
        TriggC p_contacto_165{302},p_contacto_165{303},Vel_Proceso,triggContactoCir,Z_Proceso,Prototipo_JSDaleman\WObj:=WO_Pastel;
        Mover_a_vacio;
        TriggL p_contacto_165{304},Vel_Acercamiento,triggContacto,Z_Acercamiento,Prototipo_JSDaleman\WObj:=WO_Pastel;
        Path_vacio_ejecucion p_vacio_165, 60, WO_Pastel, FALSE;
        index_vacio_destino:=310;
        Mover_a_contacto;
        TriggL p_contacto_165{305},Vel_Acercamiento,triggContacto,Z_Acercamiento,Prototipo_JSDaleman\WObj:=WO_Pastel;
        Mover_en_contacto;
        TriggC p_contacto_165{306},p_contacto_165{307},Vel_Proceso,triggContactoCir,Z_Proceso,Prototipo_JSDaleman\WObj:=WO_Pastel;
        TriggL p_contacto_165{308},Vel_Proceso,triggContacto,Z_Proceso,Prototipo_JSDaleman\WObj:=WO_Pastel;
        TriggL p_contacto_165{309},Vel_Proceso,triggContacto,Z_Proceso,Prototipo_JSDaleman\WObj:=WO_Pastel;
        Mover_a_vacio;
        TriggL p_contacto_165{310},Vel_Acercamiento,triggContacto,Z_Acercamiento,Prototipo_JSDaleman\WObj:=WO_Pastel;
        Path_vacio_ejecucion p_vacio_165, 61, WO_Pastel, FALSE;
        index_vacio_destino:=319;
        Mover_a_contacto;
        TriggL p_contacto_165{311},Vel_Acercamiento,triggContacto,Z_Acercamiento,Prototipo_JSDaleman\WObj:=WO_Pastel;
        Mover_en_contacto;
        TriggC p_contacto_165{312},p_contacto_165{313},Vel_Proceso,triggContactoCir,Z_Proceso,Prototipo_JSDaleman\WObj:=WO_Pastel;
        TriggL p_contacto_165{314},Vel_Proceso,triggContacto,Z_Proceso,Prototipo_JSDaleman\WObj:=WO_Pastel;
        TriggC p_contacto_165{315},p_contacto_165{316},Vel_Proceso,triggContactoCir,Z_Proceso,Prototipo_JSDaleman\WObj:=WO_Pastel;
        TriggC p_contacto_165{317},p_contacto_165{318},Vel_Proceso,triggContactoCir,Z_Proceso,Prototipo_JSDaleman\WObj:=WO_Pastel;
        Mover_a_vacio;
        TriggL p_contacto_165{319},Vel_Acercamiento,triggContacto,Z_Acercamiento,Prototipo_JSDaleman\WObj:=WO_Pastel;
    ENDPROC

ENDMODULE
